(* IEC 61131-3 sources: daoli-st-library/DL_Algo (part 17) *)

(* ---- FB_DL_OptimalStartStop.st ---- *)
(*
  ==================================================================
  组件名 Component  : FB_DL_OptimalStartStop
  分类   Category   : DL_Algo
  复杂度 Complexity  : cx5
  版本   Version    : 1.0.0
  功能   Purpose    : 最优启停预调度。按建筑热惯性差值提前启动：占用前依据
                      室内外温差与设定差预测恢复时长（_learned 系数在线修正
                      ——上一恢复周期实测对预测的比值按学习增益钳位推进），
                      依预测提前量给出预启动建议；占用期给出预停止建议。
                      与 EnergySavingMode 空闲节能分工互引。
  来源   Source     : t1-oscat-building（HVAC optimal start 公开语义）
  溯源   Origin     : IEC 61131-3 标准语义的道莅防御性实现；optimal start
                      预测恢复为公开暖通空调节能语义，clean-room 自研实现，
                      未复制 OSCAT 或任何厂商私有库源码。
  平台   Platform   : 纯 IEC 61131-3（Standard.library: R_TRIG，无私有库）
  分工声明 Split     : 与 FB_DL_NightPurgeSeq 分工——后者利用夜间冷量做无源
                      预冷顺控，本件为有源 HVAC 启停时刻预测调度；与存量
                      EnergySavingMode 分工——后者做占用空闲期设备降级节能，
                      本件只做启停时刻预测建议，不执行任何设备命令。
  作者   Author     : 道莅代码库 · PLC 编程专家（R58）
  ------------------------------------------------------------------
  边界 Boundary     :
                      一 代理量三句声明（R95）：fScanPeriodMin 为每次调用的
                         代表时长（代理值）；覆盖任务周期 0.1..10 分钟的调
                         用节拍；覆盖不到的区间（调用节拍外事件）由调用方
                         的占用信号沿精度兜尾；
                      二 学习系数域 [0.5..2.0]（无量纲比），越域钳定（两级
                         回退 FB32-3：先回默认 1.0，再按域钳定），学习仅在
                         bLearnEn 且恢复周期完整（启动建议发出 → 占用沿到
                         达）时推进；
                      三 预启动建议判据：占用前且预测恢复时长 ≥ 实际提前
                         余量（由剩余时间折算）——本件不接实时时钟，余量由
                         调用方经 fLeadTimeMin 传入 [分钟]；
                      四 三温度引脚（室内 / 室外 / 设定）非有限即冻结建议
                         输出为 FALSE 并置域闸故障锁存（解除 = bReset 沿）；
                      五 无全局变量、无外部变量声明、无物理地址寻址。
  修订记录 Revision  :
    2026-11-21  v1.0.0  R58 首版（批 3 · 序号 9）
  ==================================================================
*)

FUNCTION_BLOCK FB_DL_OptimalStartStop
VAR_INPUT
    bEnable       : BOOL := TRUE;   // 使能，失能建议输出安全侧 FALSE [-] / enable, disabling clears the advice
    bReset        : BOOL := FALSE;  // 复位上升沿清故障锁存与学习累计 [-] / reset rising edge clears the latch and the learning
    bOccupied     : BOOL := FALSE;  // 占用信号电平 [-] / the occupancy level
    bLearnEn      : BOOL := TRUE;   // 学习使能 [-] / the learning enable
    fTinC         : LREAL := 20.0;  // 室内温度实测 [摄氏度] / the indoor temperature [degree celsius]
    fToutC        : LREAL := 5.0;   // 室外温度实测 [摄氏度] / the outdoor temperature [degree celsius]
    fTsetC        : LREAL := 22.0;  // 占用期设定温度 [摄氏度] / the occupied setpoint [degree celsius]
    fLeadTimeMin  : LREAL := 30.0;  // 调用方传入的提前余量 [分钟] / the lead time margin fed by the caller [minute]
    fScanPeriodMin: LREAL := 1.0;   // 每次调用的代表时长 [分钟]（代理量，边界一）/ the representative duration per call [minute]
    fOptCoef      : LREAL := 4.0;   // 基础恢复系数 [分钟每开尔文每开尔文温差] / the base recovery coefficient [minute per kelvin per kelvin]
    fLearnGain    : LREAL := 0.2;   // 学习增益 [无量纲]，域 0..0.5 / the learning gain, zero through point five
END_VAR
VAR_OUTPUT
    bPreStartAdvise  : BOOL := FALSE; // 预启动建议出口 [-] / the pre start advice outlet
    bPreStopAdvise   : BOOL := FALSE; // 预停止建议出口 [-] / the pre stop advice outlet
    fPredRecoveryMin : LREAL := 0.0;  // 预测恢复时长出口 [分钟] / the predicted recovery duration outlet [minute]
    fLearnedK        : LREAL := 1.0;  // 在线学习系数出口 [无量纲] / the learned coefficient outlet, dimensionless
    bError           : BOOL := FALSE; // 域闸故障锁存标志 [-] / the domain gate fault latch flag
END_VAR
VAR
    rtOccUp  : R_TRIG; // 占用上升沿检测，段 0 无条件刷新 / the occupancy rising edge
    rtReset  : R_TRIG; // 复位沿检测，段 0 无条件刷新 / the reset edge
    _bInit   : BOOL := FALSE; // 首扫初始化完成标志（R310）/ the first scan flag
    _bLatch  : BOOL := FALSE; // 域闸故障锁存位 [-] / the domain gate latch bit
    _bRecRun : BOOL := FALSE; // 恢复期计时进行中（建议发出 → 占用沿）/ the recovery timing active
    _fRecAcc : LREAL := 0.0;  // 恢复期实测累计时长 [分钟] / the measured recovery duration accumulator [minute]
    _fPred   : LREAL := 0.0;  // 本恢复期预测值快照 [分钟] / the predicted value snapshot of this recovery
    _bPredOK : BOOL := FALSE; // 预测快照有效（学习推进前置）[-] / the prediction snapshot valid
END_VAR
VAR CONSTANT
    DL_OSS_KMIN : LREAL := 0.5; // 学习系数域下界 [无量纲] / the learned coefficient floor
    DL_OSS_KMAX : LREAL := 2.0; // 学习系数域上界 [无量纲] / the learned coefficient ceiling
    DL_OSS_GMAX : LREAL := 0.5; // 学习增益域上界 [无量纲] / the learning gain ceiling
END_VAR

// 段 0｜沿检测无条件周期刷新（禁入分支）/ segment 0, the unconditional refresh
rtOccUp(CLK := bOccupied); // 占用沿 / the occupancy edge
rtReset(CLK := bReset); // 复位沿 / the reset edge

// 段 1｜首扫初始化（R310）：学习系数回默认域内点 / segment 1, the first scan init
IF NOT _bInit THEN // 首扫一拍 / the first scan
    _bInit := TRUE; // 置首扫标志 / raise the flag
    fLearnedK := 1.0; // 学习系数回默认（FB32-3 一级回退值）/ the coefficient to the default
END_IF

// 段 2｜复位沿作用域：清故障锁存 / 清学习累计与恢复期快照 / 清建议出口（三项逐项声明）/ segment 2, the reset edge scope
IF rtReset.Q THEN // 复位沿 / the reset edge
    _bLatch := FALSE; // 作用域一：清域闸锁存 / scope one, clear the latch
    _fRecAcc := 0.0; // 作用域二：清恢复累计 / scope two, clear the recovery accumulator
    _fPred := 0.0; // 作用域二：清预测快照 / scope two, clear the prediction snapshot
    _bPredOK := FALSE; // 作用域二：清快照有效 / scope two, clear the snapshot valid
    _bRecRun := FALSE; // 作用域二：清恢复期计时 / scope two, clear the recovery timing
    bPreStartAdvise := FALSE; // 作用域三：清建议出口 / scope three, clear the advice
    bPreStopAdvise := FALSE; // 作用域三：清建议出口 / scope three, clear the advice
END_IF

// 段 3｜输入域闸（R151 全覆盖：三温度 + 系数 + 代理周期非有限与域判定，边界四）/ segment 3, the input domain gate
IF (fTinC <> fTinC) OR ((fTinC - fTinC) <> (fTinC - fTinC)) // 室内非有限 / a non finite indoor
OR (fToutC <> fToutC) OR ((fToutC - fToutC) <> (fToutC - fToutC)) // 室外非有限 / a non finite outdoor
OR (fTsetC <> fTsetC) OR ((fTsetC - fTsetC) <> (fTsetC - fTsetC)) // 设定非有限 / a non finite setpoint
OR (fScanPeriodMin <> fScanPeriodMin) OR ((fScanPeriodMin - fScanPeriodMin) <> (fScanPeriodMin - fScanPeriodMin)) // 代理周期非有限 / a non finite period
OR (fScanPeriodMin <= 0.0) // 代理周期域（≤0 无法累计）/ the period domain
OR (fLeadTimeMin <> fLeadTimeMin) OR ((fLeadTimeMin - fLeadTimeMin) <> (fLeadTimeMin - fLeadTimeMin)) // 余量非有限 / a non finite margin
OR (fOptCoef <> fOptCoef) OR ((fOptCoef - fOptCoef) <> (fOptCoef - fOptCoef)) // 系数非有限 / a non finite coefficient
OR (fOptCoef <= 0.0) // 系数域 / the coefficient domain
THEN // 任一命中 / any hit
    IF NOT _bLatch THEN // 未锁存才置位（锁存回放 R152，解除 = bReset 沿）/ latch only while unlatched
        _bLatch := TRUE; // 置域闸锁存 / raise the latch
    END_IF
END_IF
bError := _bLatch OR (fLearnGain < 0.0) OR (fLearnGain > DL_OSS_GMAX); // 故障标志聚合（锁存项 OR 增益域项，R191 名实双出口）/ the flag aggregation

// 段 4｜预测恢复时长（热惯性差值式：设定差 × 内外差因子 × 学习系数）/ segment 4, the predicted recovery
IF (NOT _bLatch) AND bEnable THEN // 域内且使能才预测 / predict only inside the domain and enabled
    IF fTinC < fTsetC THEN // 需升温场景（采暖恢复）/ a warming scenario
        fPredRecoveryMin := fOptCoef * fLearnedK * (fTsetC - fTinC) * ((fTsetC - fToutC) / (fTinC - fToutC + 20.0)); // 差值因子式（除子恒 ≥20，已证无除零）/ the delta factor form, the divisor proven at least twenty
    ELSE // 已达标或超温：恢复时长为零 / already met, the recovery zero
        fPredRecoveryMin := 0.0; // 预测零 / the prediction zero
    END_IF
ELSE // 域闸锁存或失能：预测出口清零（安全侧）/ latched or disabled, the outlet cleared
    fPredRecoveryMin := 0.0; // 清零 / cleared
END_IF

// 段 5｜学习推进（恢复周期闭合沿：占用上升沿结算，边界二）/ segment 5, the learning settlement
IF _bRecRun THEN // 恢复期计时中 / while timing the recovery
    _fRecAcc := _fRecAcc + fScanPeriodMin; // 实测累计推进（代理量，边界一）/ advance the measured accumulator
END_IF
IF rtOccUp.Q AND _bPredOK THEN // 占用沿且预测快照有效：结算学习 / the occupation edge with a valid snapshot
    _bRecRun := FALSE; // 恢复期闭合 / close the recovery
    IF (_fPred > 0.0) AND (_fRecAcc > 0.0) AND bLearnEn AND (NOT _bLatch) THEN // 四前置才推进 / the four preconditions
        IF fLearnGain > DL_OSS_GMAX THEN // 增益越域钳定（FB32-3 二级）/ the gain clamped
            fLearnGain := DL_OSS_GMAX; // 钳到上界 / clamp to the ceiling
        END_IF
        IF fLearnGain < 0.0 THEN // 增益负值钳零 / the negative gain clamped to zero
            fLearnGain := 0.0; // 钳到零 / clamp to zero
        END_IF
        fLearnedK := fLearnedK + fLearnGain * ((_fRecAcc / _fPred) - 1.0); // 比值误差推进（除子 _fPred 已证 >0）/ advance by the ratio error
        IF fLearnedK < DL_OSS_KMIN THEN // 学习系数域钳定（边界二）/ the coefficient clamped
            fLearnedK := DL_OSS_KMIN; // 钳到下界 / clamp to the floor
        ELSIF fLearnedK > DL_OSS_KMAX THEN // 越上界 / above the ceiling
            fLearnedK := DL_OSS_KMAX; // 钳到上界 / clamp to the ceiling
        END_IF
    END_IF
    _bPredOK := FALSE; // 快照消费 / consume the snapshot
    _fRecAcc := 0.0; // 累计清零备下一周期 / clear the accumulator
END_IF

// 段 6｜建议出口（边界三：不接时钟，余量由调用方传入）/ segment 6, the advice outlets
IF (NOT _bLatch) AND bEnable AND (NOT bOccupied) THEN // 占用前建议评估 / the advice before occupancy
    IF _fPred = 0.0 THEN // 本周期尚无快照（首个占用前周期）——发建议同时落快照 / no snapshot yet, raise and snapshot
        _fPred := fPredRecoveryMin; // 落预测快照 / snapshot the prediction
        _bPredOK := fPredRecoveryMin > 0.0; // 快照有效性 / the snapshot validity
        _bRecRun := fPredRecoveryMin > 0.0; // 启动恢复期计时 / start the recovery timing
    END_IF
    bPreStartAdvise := (_fPred >= fLeadTimeMin); // 预测恢复时长 ≥ 提前余量才建议 / advise when the prediction covers the margin
ELSE // 占用期或域外：预启动建议清除 / during occupancy or outside the domain
    bPreStartAdvise := FALSE; // 建议清除 / the advice cleared
END_IF
bPreStopAdvise := (NOT _bLatch) AND bEnable AND bOccupied AND (fTinC >= fTsetC); // 占用期达标预停止建议 / the pre stop advice when met during occupancy
END_FUNCTION_BLOCK

(* ---- FB_DL_OutlierFilter.st ---- *)
(*
  ==================================================================
  组件名 Component  : FB_DL_OutlierFilter
  分类   Category   : DL_Algo
  前缀   Naming     : FB_DL_ ｜ b/n/u/f/t/e/st 类型前缀制（R265）
  码位   Code ID    : 16#0002_373F / 3742（故障级）｜ 16#0002_3740 / 3741（信息级）
  版本   Version    : 1.0.0
  复杂度 Complexity  : 中
  功能   Purpose    : MAD 野点剔除滤波器：滑窗中值 + 绝对偏差中值（MAD）判野点，
                      野点丢弃并保持上次有效输出；真阶跃按连续剔除计数重基线，
                      禁「持续阶跃被永久拒绝」死锁。
  开源溯源 Origin    : 公开公式 clean-room，参考公开稳健统计教材的中值绝对偏差
                      （MAD）判据与 1.4826 正态一致性因子（分类与公式借鉴，零代码
                      复制），本件实现、闸门与码位 100% 自有。
  许可证 License    : MIT
  参考   Reference  : IEC 61131-3:2013 §6.6 算术运算符；MAD = median(|x − median|)
                      × 1.4826 公开稳健统计定义
  平台   Platform   : 纯 IEC 61131-3（FOR / 四则 / TON / 委托），三平台通用
  依赖   Depends    : FC_DL_SortIndexLReal（索引排序属主，本件双次委托，R140 /
                      R295 双承接）；Standard.library（TON）
  分工声明 Split     : FB_DL_MedianFilter（输出 = 中值，无判据）/ FB_DL_Signal
                      FrozenDetect（不变性监视）/ FB_DL_SensorDriftBaseline
                      （基线漂移）互引；本件为单点野点剔除 + 保持（R216）。
  归属 Ownership     : 本件无 TYPE 声明；全部引脚为 IEC 标准原生类型。
                      委托件码位随其属主回传（R66）。
  ------------------------------------------------------------------
  边界 Boundary     :
                      一 委托双承接（R295）：两次排序委托的返回值与 bValid 均由独立
                         变量承接后合取；委托码随属主回传（R66）；
                      二 窗长固定容量 64（禁动态分配）；nWinLen 越域钳位 + 信息级
                         3740，变更沿全窗清零（防新旧窗样本混算）；
                      三 判据 ABS(fIn − fMedian) > fNSigma × fSigmaHat + 1.0E-9 →
                         野点：不入窗、fOut 保持上次有效、bHold = TRUE、nReject + 1；
                      四 真阶跃处置（写死）：连续剔除计数 _nRejectRun ≥ nWinLen/2 →
                         判「真实阶跃」，清窗 + fIn 入窗直通 + 信息级 3741（禁死锁）；
                      五 tHoldMax 到时仍保持 → 故障级 3742 + bValid = FALSE（测点
                         疑似坏）；tonHold 段 0 无条件刷新，IN 串组态闸与保持态
                         （FB50-1 监视门控）；故障码逐拍重算不锁存（无 bReset 引脚，
                         R152 解除路径自证 = 修正组态 / 测点恢复入窗，恒可达）；
                      六 非有限 fIn → 视同野点丢弃（计数单列局部 nNonFinite，
                         不外显，不推进 _nRejectRun——测点坏与真阶跃不混淆）；
                      七 fNSigma 域闸 (0, 10] 且 tHoldMax > T#0S：非法 → 组态码
                         373F + 三件套 + RETURN 结构早退；
                      八 bEnable = FALSE 的语义写死（FB33-4 声明行）：输出冻结 +
                         窗保留（纯监视件），bHold 复位；
                      九 首拍 _bInit 全量初始化 + 首样本直通；中值 / MAD 为序不变量，
                         环形窗活样本恒为下标 0.._nFill−1（写头仅在达 _nUse 时回卷）；
                      十 无全局、无外部变量、无物理地址、无指针。
  错误码 Codes      :
    16#0002_373F【故障级】组态非法（fNSigma ≤ 0 / > 10 / 非有限，或 tHoldMax ≤ 0）
    16#0002_3740【信息级】nWinLen 越域已钳位（合法 4..64，不置 bError）
    16#0002_3741【信息级】真阶跃重基线触发（连续剔除达窗长一半，不置 bError）
    16#0002_3742【故障级】野点保持超 tHoldMax，测点疑似坏（bValid = FALSE）
  码位反证 Note     :
    373F / 3742 不可合并：373F 与窗内容无关（组态即刻判），3742 需窗已建立且持续
    保持，处置人不同（组态工程师 / 仪表工），可由 bHold 与窗状态还原（R90）；
    3740 / 3741 为信息级与故障级分属不同子带（R75 子带纪律），不可跨用。
  验收 Acceptance   :
    算法已证（脚本）：未跑 ｜ 编译器已证（三平台）：未跑
    V1 平稳序列 + 单点尖峰（10×σ）→ 剔除、fOut 保持、bHold 单拍
    V2 尖峰后立即回落 → 窗无污染；V3 真阶跃 → 连续剔除达窗长/2 后重基线直通 + 3741
    V4 fNSigma = 0 → 码 373F 早退；V5 保持超 tHoldMax → 3742 + bValid = FALSE
    V6 nWinLen = 3 → 钳 4 + 3740；V7 nWinLen 变更沿清窗；V8 首拍直通
  修订记录 Revision  :
    2026-11-21  v1.0.0  R63 首版（批 2 · 序号 7）
  ==================================================================
*)
FUNCTION_BLOCK FB_DL_OutlierFilter
VAR_INPUT
    bEnable  : BOOL := TRUE;   // 使能，FALSE 时输出冻结 + 窗保留（边界八）/ the enable, false freezes the output and keeps the window
    fIn      : LREAL := 0.0;   // 输入量 [工程单位]，必须有限 / the input value, must be finite
    nWinLen  : DINT := 16;     // 窗长 [个]，合法域 4..64，变更沿清窗 / the window length, legal four to sixty four, a change clears the window
    fNSigma  : LREAL := 4.0;   // MAD 倍数 [−]，域 (0, 10] / the MAD multiple inside the half open domain
    tHoldMax : TIME := T#5S;   // 野点连续保持上限 [毫秒]，超时判测点坏 / the hold ceiling before the point is declared broken
END_VAR
VAR_OUTPUT
    fOut     : LREAL := 0.0;            // 滤波输出 [工程单位] / the filtered output
    nReject  : UDINT := 0;             // 累计剔除计数 [个] / the accumulated reject count
    bHold    : BOOL := FALSE;          // 本拍处于保持态 [-] / the hold state of this scan
    bValid   : BOOL := FALSE;          // 输出可用 [-] / the output is usable
    eErr     : UDINT := 16#0000_0000;  // 错误码，0 = 正常 / the error code, zero is ok
    bError   : BOOL := FALSE;          // 故障标志（故障级码同拍置位，R45 配对）/ the fault flag raised with a fault level code
END_VAR
VAR
    _bInit     : BOOL := FALSE;               // 首拍初始化标志（R310 / FB50-2）/ the first scan flag
    _bHasSamp  : BOOL := FALSE;               // 已收首样本标志（首拍直通用）/ the first sample received flag
    _afWin     : ARRAY[0..63] OF LREAL;       // 采样环形窗 [工程单位]，固定容量 64 / the fixed capacity ring of samples
    _afSort    : ARRAY[0..255] OF LREAL;      // 中值排序工作数组 [工程单位] / the median sort work array
    _afDev     : ARRAY[0..255] OF LREAL;      // MAD 偏差序列工作数组 [工程单位] / the MAD deviation work array
    _aIdxM     : ARRAY[0..255] OF DINT;       // 中值排序索引承接 [下标] / the median sort index holder
    _aIdxD     : ARRAY[0..255] OF DINT;       // MAD 排序索引承接 [下标] / the MAD sort index holder
    _nHead     : DINT := 0;                   // 环形窗写头 [下标] / the ring write head
    _nFill     : DINT := 0;                   // 环形窗填充计数 [个] / the ring filled count
    _nUse      : DINT := 16;                  // 钳位后的窗长 [个] / the clamped window length
    _nUsePrev  : DINT := 0;                   // 上拍窗长快照 [个]，置 0 使首拍必触发清窗 / the previous length, zero forces one clear
    _nClrIdx   : DINT := 0;                   // 清窗遍历索引 [下标] / the clearing traversal index
    _nCopyIdx  : DINT := 0;                   // 拷贝遍历索引 [下标] / the copying traversal index
    _nMidIdx   : DINT := 0;                   // 中值下标 [下标] / the median index
    _nRejectRun: DINT := 0;                   // 连续剔除计数 [个]（真阶跃判据）/ the consecutive reject count for the step test
    _nNonFinite: DINT := 0;                   // 非有限丢弃计数 [个]（仅局部留档，不外显，R62-D7 口径）/ the dropped non finite count, local only and never exposed
    _fMedian   : LREAL := 0.0;                // 窗内中值 [工程单位] / the window median
    _fMad      : LREAL := 0.0;                // 绝对偏差中值 [工程单位] / the median absolute deviation
    _fSigmaHat : LREAL := 0.0;                // 稳健标准差估计 [工程单位] / the robust sigma estimate
    _fDev      : LREAL := 0.0;                // 本拍样本绝对偏差 [工程单位] / the absolute deviation of this scan
    _fOutLast  : LREAL := 0.0;                // 最近一次有效输出（保持源）[工程单位] / the last valid output used while holding
    _bHoldActive : BOOL := FALSE;             // 保持态寄存器（跨拍保持，tonHold 驱动源）/ the hold state register driving the timer
    _bCfgBad   : BOOL := FALSE;               // 组态非法标记（逐拍重算）/ the configuration fault flag
    _bWinClamp : BOOL := FALSE;               // 窗长钳位标记（逐拍重算，信息级 3740）/ the window clamp flag
    _bStepReb  : BOOL := FALSE;               // 真阶跃重基线标记（逐拍重算，信息级 3741）/ the step rebuild flag
    _bHoldOut  : BOOL := FALSE;               // 本拍保持出口位（统一出口映射）/ the hold outlet bit of this scan
    _bRejectI  : BOOL := FALSE;               // 本拍拒绝内部位 / the internal reject bit of this scan
    _bFinIn    : BOOL := FALSE;               // 输入有限闸结果（逐拍重算）/ the input finiteness gate result
    _bFinSig   : BOOL := FALSE;               // fNSigma 有限闸结果（逐拍重算）/ the sigma pin finiteness gate result
    _bSortRet  : BOOL := FALSE;               // 中值委托返回值承接量（独立承接，R295）/ the median delegate return holder
    _bSortValid: BOOL := FALSE;               // 中值委托可用位承接量 / the median delegate valid holder
    _bSortRet2 : BOOL := FALSE;               // MAD 委托返回值承接量（独立承接，R295）/ the MAD delegate return holder
    _bSortValid2: BOOL := FALSE;              // MAD 委托可用位承接量 / the MAD delegate valid holder
    _uSortErr  : UDINT := 16#0000_0000;       // 中值委托码承接量 [码] / the median delegate code holder
    _uSortErr2 : UDINT := 16#0000_0000;       // MAD 委托码承接量 [码] / the MAD delegate code holder
    _bSortErr  : BOOL := FALSE;               // 中值委托故障位承接量 / the median delegate fault holder
    _bSortErr2 : BOOL := FALSE;               // MAD 委托故障位承接量 / the MAD delegate fault holder
    tonHold    : TON;                         // 保持超时定时器，段 0 无条件刷新 / the hold timeout timer refreshed unconditionally
END_VAR  // R64 结构补齐：VAR 段缺失的 END_VAR（门禁机械修复）
VAR CONSTANT
    DL_OF_WMAX  : DINT := 64;       // 窗容量上界 [个]，与数组容量一致 / the window capacity aligned with the array
    DL_OF_WMIN  : DINT := 4;        // 窗长下界 [个] / the window floor
    DL_OF_NSIGMAX : LREAL := 10.0;  // MAD 倍数上界 [−] / the MAD multiple ceiling
    DL_OF_NSIGZERO: LREAL := 0.0;   // MAD 倍数零常量 [−] / the MAD multiple zero constant
    DL_OF_MADK    : LREAL := 1.4826; // MAD 正态一致性因子 [−] / the MAD normal consistency factor
    DL_OF_EPS     : LREAL := 1.0E-9; // 判据容差 [工程单位] / the criterion tolerance
    DL_OF_STEPDIV : LREAL := 2.0;   // 真阶跃判据除子 [−]（窗长一半）/ the step criterion divisor of one half
    DL_OF_ZERO    : LREAL := 0.0;   // 实数零常量 [工程单位] / the real zero constant
    DL_OF_ONE     : DINT := 1;      // 整型一常量 [个] / the integer one constant
    DL_OF_TWO     : DINT := 2;      // 整型二常量 [个]（中值判据最少样本）/ the integer two constant, the minimum for a median
    DL_OF_ZEROI   : DINT := 0;      // 整型零常量 [个] / the integer zero constant
    DL_OF_TIME0   : TIME := T#0S;   // 时间零常量 [毫秒] / the time zero constant
END_VAR

// 段 0｜组态闸先行 + 定时器无条件周期刷新（禁入分支，R7；监视 TON 串组态闸，FB50-1）/ segment 0, the configuration gate first and the unconditional timer refresh
_bFinSig := (fNSigma = fNSigma) AND ((fNSigma - fNSigma) = (fNSigma - fNSigma)); // fNSigma 有限 / the sigma pin is finite
_bCfgBad := (NOT _bFinSig) OR (fNSigma <= DL_OF_NSIGZERO) OR (fNSigma > DL_OF_NSIGMAX) OR (tHoldMax <= DL_OF_TIME0); // 组态非法（MAD 倍数域外或保持上限非正）/ an illegal configuration
tonHold(IN := _bHoldActive AND (NOT _bCfgBad), PT := tHoldMax); // 保持超时计时（串组态闸，防复位同拍重锁，FB50-1）/ the hold timeout with the configuration gate in series

// 段 1｜首拍初始化与窗长接管预派生（FB50-2）/ segment 1, the first scan init
IF NOT _bInit THEN // 首拍一拍 / the first scan
    _bInit := TRUE; // 置首拍标志 / raise the first scan flag
    _bHasSamp := FALSE; // 首样本标志显式清零（触发直通）/ clear the first sample flag so the pass through triggers
    _nFill := DL_OF_ZEROI; // 填充计数显式清零 / clear the filled count explicitly
    _nHead := DL_OF_ZEROI; // 写头显式清零 / clear the write head explicitly
    _nUsePrev := DL_OF_ZEROI; // 窗长快照置 0，使段 2 变更沿必然触发一次清窗 / zero the snapshot so the change edge clears the window once
    _nRejectRun := DL_OF_ZEROI; // 连续剔除计数显式清零 / clear the consecutive reject count explicitly
    _nNonFinite := DL_OF_ZEROI; // 非有限计数显式清零 / clear the non finite count explicitly
    _bHoldActive := FALSE; // 保持态显式清零 / clear the hold state explicitly
    _fOutLast := DL_OF_ZERO; // 最近有效输出显式清零 / clear the last valid output explicitly
    FOR _nClrIdx := DL_OF_ZEROI TO DL_OF_WMAX - DL_OF_ONE DO // 有界遍历全容量 / the bounded traversal over the full capacity
        _afWin[_nClrIdx] := DL_OF_ZERO; // 窗元素逐项清零 / zero every window element
    END_FOR
END_IF

// 段 2｜窗长钳位与变更沿全窗清零（边界二）/ segment 2, the window length clamp and the full clear
_bWinClamp := FALSE; // 钳位标记预清零（单拍信息位，段 8 统一映射）/ preset the clamp flag false
_bStepReb := FALSE; // 重基线标记预清零（单拍信息位）/ preset the rebuild flag false
_bHoldOut := FALSE; // 保持出口位预清零（单拍信息位，R256 统一出口预置）/ preset the hold outlet bit false
_bRejectI := FALSE; // 拒绝内部位预清零（单拍位）/ preset the reject bit false
_nUse := nWinLen; // 窗长接管 [个] / take the window length
IF (_nUse < DL_OF_WMIN) OR (_nUse > DL_OF_WMAX) THEN // 窗长越域 / the length is out of the domain
    _bWinClamp := TRUE; // 置钳位标记（信息级 3740）/ raise the clamp flag
    IF _nUse < DL_OF_WMIN THEN // 下界钳位 / the floor clamp
        _nUse := DL_OF_WMIN; // 钳到下界 [个] / clamp to the floor
    ELSE // 上界钳位 / the ceiling clamp
        _nUse := DL_OF_WMAX; // 钳到容量 [个] / clamp to the capacity
    END_IF
END_IF
IF _nUse <> _nUsePrev THEN // 窗长变更沿（含首拍）/ the length change edge, the first scan included
    _nHead := DL_OF_ZEROI; // 写头回零 / reset the write head
    _nFill := DL_OF_ZEROI; // 填充计数回零 / reset the filled count
    _nRejectRun := DL_OF_ZEROI; // 连续剔除计数回零 / reset the consecutive reject count
    _bHasSamp := FALSE; // 窗已清，首样本语义复位 / the window is cleared, the first sample semantics reset
    FOR _nClrIdx := DL_OF_ZEROI TO DL_OF_WMAX - DL_OF_ONE DO // 有界遍历全容量 / the bounded traversal over the full capacity
        _afWin[_nClrIdx] := DL_OF_ZERO; // 窗元素逐项清零（禁陈旧样本混算）/ zero every window element so no stale sample mixes in
    END_FOR
    _nUsePrev := _nUse; // 快照本拍窗长 / snapshot the length
END_IF

// 段 3｜失能分支：输出冻结 + 窗保留（边界八声明行）/ segment 3, the disabled branch freezes the output
IF NOT bEnable THEN // 失能 / disabled
    fOut := _fOutLast; // 冻结最后有效输出 [工程单位] / freeze the last valid output
    bHold := FALSE; // 保持态复位 / the hold state resets
    bValid := FALSE; // 失能即不可用 / the output is not usable while disabled
    bError := FALSE; // 失能不是故障 / a disabled device is not a fault
    eErr := 16#0000_0000; // 失能不发码 / no code is emitted while disabled
    _bHoldActive := FALSE; // 保持态寄存器复位（tonHold 断输入）/ clear the hold state register
    RETURN; // 早退，窗保留；nReject 为累计量按 R187 不清零（保持语义由本注释表达，禁自赋值行）/ early return with the window kept, the accumulated reject count is kept per the pulse discipline, expressed by this comment without a dead statement
END_IF

// 段 4｜组态非法结构早退（边界七，出口三件套 + RETURN）/ segment 4, the structural early exit on an illegal configuration
IF _bCfgBad THEN // 组态非法 / an illegal configuration
    fOut := _fOutLast; // 输出保持最近有效值 [工程单位] / keep the last valid output
    bHold := FALSE; // 保持态复位 / the hold state resets
    bValid := FALSE; // 输出不可用 / the output is not usable
    eErr := 16#0002_373F; // 故障级：组态非法 / fault grade, an illegal configuration
    bError := TRUE; // 同拍置故障标志（R45 配对）/ raise the fault flag on the same scan
    _bHoldActive := FALSE; // 保持态寄存器复位 / clear the hold state register
    RETURN; // 早退，判据段不可达 / early return, the criterion segment is unreachable
END_IF

// 段 5｜输入有限闸（边界六）/ segment 5, the input finiteness gate
_bFinIn := (fIn = fIn) AND ((fIn - fIn) = (fIn - fIn)); // 输入有限 / the input is finite
IF NOT _bHasSamp THEN // 首样本直通（边界十）/ the first sample passes straight through
    _afWin[_nHead] := fIn; // 首样本入窗 [工程单位] / the first sample enters the window
    _nHead := _nHead + DL_OF_ONE; // 写头推进 / advance the head
    IF _nHead >= _nUse THEN // 回卷 / wrap
        _nHead := DL_OF_ZEROI; // 写头回零 / reset the head
    END_IF
    _nFill := _nFill + DL_OF_ONE; // 填充计数推进 [个] / advance the filled count
    fOut := fIn; // 首拍直通 [工程单位] / the first scan passes straight through
    _fOutLast := fIn; // 有效输出快照 [工程单位] / snapshot the valid output
    _bHasSamp := TRUE; // 置首样本标志 / raise the first sample flag
    bHold := FALSE; // 无保持 / no hold
    bValid := TRUE; // 输出可用 / the output is usable
    eErr := 16#0000_0000; // 正常 / ok
    bError := FALSE; // 无故障 / no fault
    RETURN; // 早退 / early return
END_IF

// 段 6｜非有限输入：视同野点丢弃（边界六，计数单列，不推进连续剔除计数）/ segment 6, a non finite input is dropped like an outlier
IF NOT _bFinIn THEN // 输入坏 / the input is broken
    _nNonFinite := _nNonFinite + DL_OF_ONE; // 非有限计数推进（仅局部留档）/ advance the non finite count, local only
    _bHoldActive := TRUE; // 置保持态（tonHold 持续计时）/ raise the hold state
    fOut := _fOutLast; // 输出保持 [工程单位] / keep the output
    bHold := TRUE; // 保持出口位 / the hold outlet
    bValid := TRUE; // 保持值本身可用（未超时前）/ the held value is still usable before the timeout
    eErr := 16#0000_0000; // 信息级不占故障位 / no fault code for a single drop
    bError := FALSE; // 无故障 / no fault
    RETURN; // 早退 / early return
END_IF

// 段 7｜中值与 MAD 计算（两次委托，双承接 R295；活样本恒为 0.._nFill−1，边界九）/ segment 7, the median and the MAD via two delegates
IF _nFill >= DL_OF_TWO THEN // 窗内至少两样本才建判据（单样本无离散度语义）/ the criterion needs at least two samples
    FOR _nCopyIdx := DL_OF_ZEROI TO _nFill - DL_OF_ONE DO // 有界遍历活样本（上界已证 ≤ 64）/ the bounded traversal over the live samples
        _afSort[_nCopyIdx] := _afWin[_nCopyIdx]; // 拷贝到排序工作数组 [工程单位] / copy into the sort work array
    END_FOR
    _bSortRet := FC_DL_SortIndexLReal(afValues := _afSort, nCount := _nFill, aIdx => _aIdxM, bValid => _bSortValid, eErr => _uSortErr, bError => _bSortErr); // 中值排序委托 / delegate the median sort
    _nMidIdx := (_nFill - DL_OF_ONE) / DL_OF_TWO; // 中值下标（偶数窗取下中值）[下标] / the median index, the lower median for an even window
    _fMedian := _afSort[_aIdxM[_nMidIdx]]; // 窗内中值 [工程单位] / the window median
    FOR _nCopyIdx := DL_OF_ZEROI TO _nFill - DL_OF_ONE DO // 有界遍历活样本 / the bounded traversal over the live samples
        _afDev[_nCopyIdx] := ABS(_afWin[_nCopyIdx] - _fMedian); // 绝对偏差序列 [工程单位] / the absolute deviation series
    END_FOR
    _bSortRet2 := FC_DL_SortIndexLReal(afValues := _afDev, nCount := _nFill, aIdx => _aIdxD, bValid => _bSortValid2, eErr => _uSortErr2, bError => _bSortErr2); // MAD 排序委托（双承接）/ delegate the MAD sort with the dual catch
    _fMad := _afDev[_aIdxD[_nMidIdx]]; // 绝对偏差中值 [工程单位] / the median absolute deviation
    _fSigmaHat := _fMad * DL_OF_MADK; // 稳健标准差估计 [工程单位] / the robust sigma estimate
    IF (NOT (_bSortRet AND _bSortValid)) OR _bSortErr OR (NOT (_bSortRet2 AND _bSortValid2)) OR _bSortErr2 THEN // 任一委托失败（双承接合取，R295）/ either delegate failed under the dual catch
        fOut := _fOutLast; // 输出保持 [工程单位] / keep the output
        bHold := FALSE; // 保持态不置（委托失败非野点）/ the hold is not raised, a delegate failure is not an outlier
        bValid := FALSE; // 输出不可用 / the output is not usable
        eErr := _uSortErr; // 委托码回传（码随属主，R66）/ replay the delegate code
        bError := _bSortErr OR _bSortErr2; // 委托故障位回传 / replay the delegate fault bits
        RETURN; // 早退 / early return
    END_IF
ELSE // 窗内样本不足：判据挂起，直接接受本拍样本 / too few samples, the criterion suspends and the sample is accepted
    _fMedian := _afWin[DL_OF_ZEROI]; // 中值占位（不参与判据）[工程单位] / a placeholder median, not used by the criterion
    _fSigmaHat := DL_OF_ZERO; // 离散度占位零 [工程单位] / a placeholder sigma of zero
END_IF

// 段 8｜野点判据与真阶跃处置（边界三四；本拍接受语义优先于超时迁移，R275）/ segment 8, the outlier criterion and the true step handling
_fDev := ABS(fIn - _fMedian); // 本拍绝对偏差 [工程单位] / the absolute deviation of this scan
IF _nFill >= DL_OF_TWO THEN // 判据已建立才比较 / the comparison runs only with a built criterion
    IF _fDev > (fNSigma * _fSigmaHat) + DL_OF_EPS THEN // 超出 MAD 带外：疑似野点 / beyond the MAD band, a suspected outlier
        _nRejectRun := _nRejectRun + DL_OF_ONE; // 连续剔除计数推进 [个] / advance the consecutive reject count
        IF DINT_TO_LREAL(_nRejectRun) >= (DINT_TO_LREAL(_nUse) / DL_OF_STEPDIV) THEN // 连续剔除达窗长一半：判真阶跃（边界四，禁死锁）/ the consecutive rejects reach half the window, a true step
            _nHead := DL_OF_ZEROI; // 清窗：写头回零 / the rebuild, the head resets
            _nFill := DL_OF_ONE; // 填充计数重置为新基线首样本 [个] / the fill resets to the first sample of the new base
            _nRejectRun := DL_OF_ZEROI; // 连续剔除计数清零 / clear the consecutive reject count
            FOR _nClrIdx := DL_OF_ZEROI TO DL_OF_WMAX - DL_OF_ONE DO // 有界遍历全容量 / the bounded traversal over the full capacity
                _afWin[_nClrIdx] := DL_OF_ZERO; // 窗元素逐项清零 / zero every window element
            END_FOR
            _afWin[DL_OF_ZEROI] := fIn; // 新基线首样本入窗 [工程单位] / the new base sample enters the window
            _nHead := DL_OF_ONE; // 写头推进一位 / advance the head by one
            fOut := fIn; // 阶跃直通 [工程单位] / the step passes straight through
            _fOutLast := fIn; // 有效输出快照 [工程单位] / snapshot the valid output
            _bStepReb := TRUE; // 置重基线标记（信息级 3741）/ raise the rebuild flag
            _bHoldActive := FALSE; // 保持态解除 / release the hold state
            bHold := FALSE; // 保持出口位复位 / the hold outlet resets
            bValid := TRUE; // 输出可用 / the output is usable
            bError := FALSE; // 信息级不置故障位 / the informational code never raises the fault bit
            IF _bWinClamp THEN // 同拍窗长钳位（信息级优先序：钳位先于重基线）/ a clamp on the same scan
                eErr := 16#0002_3740; // 信息级：窗长越域已钳位 / informational, the length was clamped
            ELSE // 无钳位 / no clamp
                eErr := 16#0002_3741; // 信息级：真阶跃重基线触发 / informational, a true step rebuilt the base
            END_IF
            RETURN; // 早退 / early return
        ELSE // 单点野点：丢弃并保持（边界三）/ a single outlier, dropped with the output held
            _bHoldActive := TRUE; // 置保持态 / raise the hold state
            _bHoldOut := TRUE; // 保持出口位置位（段 10 映射）/ raise the hold outlet bit
            _bRejectI := TRUE; // 拒绝位置位 / raise the reject bit
            fOut := _fOutLast; // 输出保持上次有效值 [工程单位] / hold the last valid output
        END_IF
    ELSE // 带内：接受样本 / inside the band, the sample is accepted
        _afWin[_nHead] := fIn; // 样本入窗 [工程单位] / the sample enters the window
        _nHead := _nHead + DL_OF_ONE; // 写头推进 / advance the head
        IF _nHead >= _nUse THEN // 回卷 / wrap
            _nHead := DL_OF_ZEROI; // 写头回零 / reset the head
        END_IF
        IF _nFill < _nUse THEN // 窗未满才累加 / count only while not full
            _nFill := _nFill + DL_OF_ONE; // 填充计数推进 [个] / advance the filled count
        END_IF
        _nRejectRun := DL_OF_ZEROI; // 连续剔除计数清零 / clear the consecutive reject count
        _bHoldActive := FALSE; // 保持态解除 / release the hold state
        fOut := fIn; // 接受直通 [工程单位] / the accepted sample passes straight through
        _fOutLast := fIn; // 有效输出快照 [工程单位] / snapshot the valid output
    END_IF
ELSE // 判据挂起拍：直接接受（窗建立期）/ the criterion suspended, the sample is accepted while the window builds
    _afWin[_nHead] := fIn; // 样本入窗 [工程单位] / the sample enters the window
    _nHead := _nHead + DL_OF_ONE; // 写头推进 / advance the head
    IF _nHead >= _nUse THEN // 回卷 / wrap
        _nHead := DL_OF_ZEROI; // 写头回零 / reset the head
    END_IF
    IF _nFill < _nUse THEN // 窗未满才累加 / count only while not full
        _nFill := _nFill + DL_OF_ONE; // 填充计数推进 [个] / advance the filled count
    END_IF
    _nRejectRun := DL_OF_ZEROI; // 连续剔除计数清零 / clear the consecutive reject count
    _bHoldActive := FALSE; // 保持态解除 / release the hold state
    fOut := fIn; // 接受直通 [工程单位] / the accepted sample passes straight through
    _fOutLast := fIn; // 有效输出快照 [工程单位] / snapshot the valid output
END_IF

// 段 9｜保持超时判据（边界五：测点疑似坏）/ segment 9, the hold timeout test
IF tonHold.Q THEN // 保持超 tonHoldMax / the hold exceeded its ceiling
    fOut := _fOutLast; // 输出保持（安全侧冻结）[工程单位] / hold the output
    bHold := TRUE; // 保持出口位 / the hold outlet
    bValid := FALSE; // 测点疑似坏，输出不可用 / the point is suspected broken, the output is unusable
    eErr := 16#0002_3742; // 故障级：保持超时 / fault grade, the hold timed out
    bError := TRUE; // 同拍置故障标志（R45 配对）/ raise the fault flag on the same scan
    RETURN; // 早退 / early return
END_IF

// 段 10｜统一出口（单拍位映射 + 累计计数单点写入，R187 / FB51-8）/ segment 10, the unified outlet
bHold := _bHoldOut; // 保持出口位（段 2 预置 + 段 8 置位映射）/ the hold outlet mapped from the preset and the raise
IF _bRejectI THEN // 本拍发生拒绝 / a reject happened on this scan
    nReject := nReject + 1; // 累计剔除计数单点写入 [个] / the accumulated reject count written at this single point
END_IF
bValid := TRUE; // 输出可用 / the output is usable
bError := FALSE; // 无故障 / no fault
IF _bWinClamp THEN // 窗长钳位（信息级，逐拍重算）/ the length clamp, informational and recomputed
    eErr := 16#0002_3740; // 信息级：窗长越域已钳位 / informational, the length was clamped
ELSE // 无事件 / no event
    eErr := 16#0000_0000; // 正常 / ok
END_IF
END_FUNCTION_BLOCK

(* ---- FB_DL_OverrideSelector.st ---- *)
(*
  FB_DL_OverrideSelector  —  高选/低选超驰选择器 / High-select and low-select override selector
  分类 Category : DL_Algo
  版本 Version  : 1.0.0
  来源 Source   : t2-5-modpid — 超驰选择族零检索深化
  溯源 Origin   : clean-room 实现，未复制任何源码行
  功能 Function : 1) 对前 nCh 路输入按 eSel 做 eHigh（高选）/ eLow（低选）仲裁，
                  输出胜出值 fOut 与胜出通道号 uWin（1 基；0 = 无有效输入）；
                  2) 只统计 aEn 使能且非有限的通道；平值取首路（严格 > / < 比较）；
                  3) nCh <= 0 或 > 8 → 故障级 03A3 拒绝；eSel 落枚举域外 → CASE ELSE → 03A4；
                  4) 首次出现有效输出沿置信息级 0489；全通道无效置信息级 048A。
  边界 Boundary : ① 判界先行：通道数域闸在仲裁前完成；
                  ② 仲裁循环带守卫计数，防失控；
                  ③ 非有限输入自动失格（NaN 自反判），不参与仲裁；
                  ④ 无 GVL 依赖：纯引脚输入输出，无外部变量引用，无物理 IO 地址。
  依赖 Depends  : 仅 Standard.library（LREAL/REAL 算术）
  码表 Error codes（Algo 段 0002，窗口 03A3~03A4 / 0489~048A）:
    16#0002_03A3 故障级：通道数非法（nCh <= 0 或 > 8），输出强制无效，bError = TRUE
    16#0002_03A4 故障级：选择模式落 CASE ELSE 兜底（非法 eSel），bError = TRUE
    16#0002_0489 信息级：首次有效输出沿（uWin 从 0 变非 0）
    16#0002_048A 信息级：全通道无效（无有效输出）
  修订历史 Revision :
    2026-11-19  v1.0.0  R41 首版（批次 2 · 序号 3）
*)

TYPE E_DL_OvrMode :
(
    eHigh := 0,    // 高选：取最大有效值 / High-select, take the maximum valid value
    eLow  := 10    // 低选：取最小有效值 / Low-select, take the minimum valid value
);
END_TYPE

FUNCTION_BLOCK FB_DL_OverrideSelector
VAR_INPUT
    aIn          : ARRAY[1..8] OF REAL;   // 候选输入数组 [EU] / Candidate inputs
    aEn          : ARRAY[1..8] OF BOOL;   // 通道使能数组 [-] / Channel enable array
    nCh          : INT := 8;          // 参与通道数 [路]，域 1..8 / Active channel count
    eSel         : E_DL_OvrMode := E_DL_OvrMode.eHigh;  // 选择模式 / Selection mode
END_VAR
VAR_OUTPUT
    fOut         : REAL;              // 胜出输出 [EU] / Winning output
    uWin         : UINT;              // 胜出通道号 [路]，0 = 无有效输入 / Winning channel, 0 = none
    bValid       : BOOL;              // 输出有效标志 / Output valid flag
    bError       : BOOL;              // 故障级标志（信息级不置位）/ Fault-level flag
    nErrId       : UDINT;             // 事件码，0 = 无事件 / Event code
END_VAR
VAR
    _uWin        : UINT;              // 内部胜出通道（出口镜像）/ Internal winning channel
    _fBest       : REAL;              // 当前最优值 [EU] / Current best value
    _bFound      : BOOL;              // 是否找到有效候选 / Valid candidate found
    _bAnyPrev    : BOOL;              // 上拍有输出口径镜像（首次有效沿判据）/ Previous valid mirror
    _nGuard      : INT;               // 仲裁守卫计数 [次] / Arbitration guard counter
    i            : INT;               // 仲裁循环游标 [索引] / Arbitration loop cursor
    _bNonFin     : BOOL;              // 当前元素非有限标志 / Non-finite flag of current element
END_VAR

(* —— 段 0｜单拍量预清零（纯派生件，无定时器/沿实例） —— *)
uWin := 0;                          // 胜出通道缺省 0（无有效输入）
fOut := 0.0;                        // 胜出值缺省 0
bValid := FALSE;                    // 有效出口缺省 FALSE
bError := FALSE;                    // 故障标志缺省 FALSE
nErrId := 16#0000_0000;             // 事件码缺省无事件
_bFound := FALSE;                   // 候选未找到
_uWin := 0;                         // 内部胜出清零
_nGuard := 0;                       // 守卫清零

(* —— 段 1｜判界先行：通道数域闸（越界直接故障出口，R101 配对） —— *)
IF (nCh <= 0) OR (nCh > 8) THEN
    nErrId := 16#0002_03A3;         // 故障级：通道数非法
    bError := TRUE;                 // 故障码配对置位
    RETURN;                         // 直接出口 / early exit
END_IF

(* —— 段 2｜仲裁：CASE 全覆盖 + ELSE 兜底落 03A4（R190：模式归因唯一） —— *)
CASE eSel OF

E_DL_OvrMode.eHigh:
    FOR i := 1 TO nCh DO
        _nGuard := _nGuard + 1;                 // 守卫递增
        IF _nGuard > 8 THEN
            EXIT;                               // 守卫兜底退出（理论不可达）
        END_IF
        _bNonFin := (aIn[i] <> aIn[i]) OR ((aIn[i] - aIn[i]) <> (aIn[i] - aIn[i]));
                                                    // NaN 自反判 OR Inf 差值自减判
        IF aEn[i] AND (NOT _bNonFin) THEN
            IF (NOT _bFound) OR (aIn[i] > _fBest) THEN
                _fBest := aIn[i];               // 高选：严格大于才换（平值取首路）
                _uWin := INT_TO_UINT(i);        // 记胜出通道
                _bFound := TRUE;                // 已找到
            END_IF
        END_IF
    END_FOR

E_DL_OvrMode.eLow:
    FOR i := 1 TO nCh DO
        _nGuard := _nGuard + 1;                 // 守卫递增
        IF _nGuard > 8 THEN
            EXIT;                               // 守卫兜底退出（理论不可达）
        END_IF
        _bNonFin := (aIn[i] <> aIn[i]) OR ((aIn[i] - aIn[i]) <> (aIn[i] - aIn[i]));
                                                    // 非有限判定同高选口径
        IF aEn[i] AND (NOT _bNonFin) THEN
            IF (NOT _bFound) OR (aIn[i] < _fBest) THEN
                _fBest := aIn[i];               // 低选：严格小于才换（平值取首路）
                _uWin := INT_TO_UINT(i);        // 记胜出通道
                _bFound := TRUE;                // 已找到
            END_IF
        END_IF
    END_FOR

ELSE
    nErrId := 16#0002_03A4;         // 故障级：非法选择模式兜底
    bError := TRUE;                 // 故障码配对置位
    RETURN;                         // 直接出口（出口保持缺省无效）/ early exit

END_CASE

(* —— 段 3｜出口单点映射（名实同源） —— *)
IF _bFound THEN
    fOut := _fBest;                 // 胜出值出口
    uWin := _uWin;                  // 胜出通道出口
    bValid := TRUE;                 // 有效出口
    IF NOT _bAnyPrev THEN
        nErrId := 16#0002_0489;     // 信息级：首次有效输出沿
    END_IF
ELSE
    uWin := 0;                      // 无有效输入（哨兵零通道）
    nErrId := 16#0002_048A;         // 信息级：全通道无效
END_IF
_bAnyPrev := _bFound;               // 首次有效沿判据快照

END_FUNCTION_BLOCK

(* ---- FB_DL_ParticleCounterStat.st ---- *)
//==============================================================================
// 功能块：FB_DL_ParticleCounterStat ｜ 中文名称：尘埃粒子计数器统计与等级判定
// 所属子库：DL_Algo ｜ 版本：v1.0.0 ｜ 兼容：CODESYS V3.5+ / TwinCAT 3 / 汇川 InoProShop
// 功能描述：6 路粒径计数（0.1/0.2/0.3/0.5/1.0/5.0 微米）→ 浓度（颗每
//           立方米）→ ISO 14644-1:2015 Table 1 等级判定（生成式 Cn =
//           10^N 乘 (0.1/D)^2.08，N 允许 0.5 步进）→ 连续 N 个采样超限
//           才报警 → 失采检测。等级判定采用 Table 1 常量表锚定 + 档内
//           LOG 对数插值：** 幂运算符跨平台不可用，改用「整数档查表
//           + LOG 对数插值」，由生成式恒等式 conc/L_N = 10^(level-N)
//           保证档内插值与公式严格一致，不引入近似误差。表内「—」
//           （无限制）格跳过不参与判定。只统计与判定，不控净化设备
//           （FFU/风淋室由上位调度，本件零执行输出）。
// 开源溯源 (Origin)：道莅原创实现（参考 ISO 14644-1:2015 Table 1 公开分级口径 分类与参数域）
// 单位表：粒子计数[颗] / 采样体积[L] / 浓度[颗/m³] / 等级[—] / 采样周期[min] / 确认数[个]
// 错误码表：16#0002_3301 信息级（采样失采，等级不可判，等级清零不沿用，
//           不置 bError）/ 16#0002_3302 信息级（等级超 9 钳 9.0，或通道
//           浓度超最深有表值档且更高档无限制被表驱动跳过，不置 bError）/
//           16#0002_3305 预留禁用（不得挪用）/ 16#0002_3310 故障级（采样
//           体积小于等于 0 或组态非法，置 bError）/ 16#0002_3311 故障级
//           （浮点输入非有限，置 bError）/ 16#0002_3312 预留禁用（不得挪用）
// 状态机：E_DL_ParticleStatState（eIdle=0 / eSampling=10 / eLost=20 /
//           eFault=99），CASE 含 ELSE 兜底，ELSE 复用 3311（§3 未为本件
//           单列兜底槽，非法状态按「数据不可信」同语义处置，不得越段
//           加码）并回 eFault、等级清零（安全侧 = 不给达标假象）
// 边界行为：① 浮点输入非有限（NaN 自反判 + Inf 幅值上限判）→ 故障 3311，
//           等级清零；② fSampleVolL 小于等于防除零下限、fClassTarget 超
//           1.0~9.0 域、nConfirmSamples 超 1~10 域、tSampleTime 非正 →
//           故障 3310，先判后除防除零；③ 全通道计数为 0 且脉冲到达 =
//           合法 0 浓度，不判失采（失采只由失采定时器时间判据裁决）；
//           ④ 失采（间隔超 2 倍采样周期）→ 信息 3301 + 等级清零 +
//           bValid := FALSE，禁止沿用旧等级（旧等级会让洁净室误报达标）；
//           bOverLimit 报警锁存保持（已确认的超限事实不因失采被掩盖，
//           恢复采样后由新数据重新裁决）；⑤ 等级超 9 → 判 9.0 并信息
//           3302；⑥ 通道浓度超该通道最深有表值档且更高档为「—」→ 该
//           通道表驱动跳过不参与判定并信息 3302（披露：跳过通道的更高
//           污染贡献不参与最严等级裁决，靠 3302 可观测提示，若全通道
//           均被跳过则等级判不可用）；⑦ 上电首拍 bValid := FALSE；
//           ⑧ 失能 → eIdle、等级清零、报警清除；⑨ 失采定时器经脉冲沿
//           「断输入一拍」重启计时，失采门槛严格等于 2 倍采样周期
//           （R40 家族）。
// 修订历史：v1.0.0 2026-11-17 首版（R25 派单 · §4.2）
//==============================================================================
(*------------------------------------------------------------------------------
 * 枚举: E_DL_ParticleStatState（归属 DL_Algo，与 FB_DL_ParticleCounterStat 同文件）
 *----------------------------------------------------------------------------*)
TYPE E_DL_ParticleStatState :
(
    eIdle     := 0,    // 失能/待机：等级输出 0，报警清零 / Idle: class zeroed, alarm cleared
    eSampling := 10,   // 采样有效：最近一次脉冲已判定，等级可用 / Sampling: last pulse judged, class usable
    eLost     := 20,   // 失采：超 2 倍采样周期无脉冲，等级不可判 / Lost: no pulse within twice the sample period
    eFault    := 99    // 故障兜底态：组态非法或非有限，等级清零 / Fault fallback: config invalid or non-finite, class zeroed
);
END_TYPE
FUNCTION_BLOCK FB_DL_ParticleCounterStat
VAR_INPUT
    auCounts        : ARRAY[0..5] OF UDINT;    // 本采样周期各粒径计数 [颗]，通道序 0.1/0.2/0.3/0.5/1.0/5.0 微米 / counts per channel [particles], channels 0.1/0.2/0.3/0.5/1.0/5.0 um
    fSampleVolL     : LREAL := 1.0;            // 采样体积 [L]，域大于 0 / Sample volume [L], domain > 0
    bSamplePulse    : BOOL;                    // 采样周期完成脉冲，上升沿取数 / Sample-complete pulse, latched on rising edge
    fClassTarget    : LREAL := 7.0;            // 目标等级 [—]，1.0~9.0，0.5 步进 / Target class, 1.0~9.0, 0.5 steps
    nConfirmSamples : INT := 3;                // 连续超限确认数 [个]，1~10 / Consecutive over-limit confirmations, 1~10
    tSampleTime     : TIME := T#1M;            // 采样周期 [min]，用于失采判定 / Sample period [min], loss detection basis
    bEnable         : BOOL;                    // 总使能 / Master enable
    bReset          : BOOL;                    // 复位，上升沿清状态与计数 / Reset, rising edge clears state and counters
END_VAR
VAR_OUTPUT
    afConcM3        : ARRAY[0..5] OF LREAL;    // 各粒径浓度 [颗/m³] / Concentration per channel [particles/m3]
    fClassMeasured  : LREAL;                   // 实测等级 [—]，0.0 = 不可判 / Measured class, 0.0 = not judgeable
    bClassOk        : BOOL;                    // 实测等级不超过目标等级 / Measured class within target
    bOverLimit      : BOOL;                    // 连续确认后的超限报警锁存 / Confirmed over-limit alarm latch
    bSampleLost     : BOOL;                    // 失采标志 / Sample-loss flag
    tSinceSample    : TIME;                    // 距上次成功采样耗时 [min] / Time since last accepted sample [min]
    uSampleCount    : UDINT;                   // 累计采样次数 [次]，饱和计数 / Cumulative sample count, saturated
    uOverCount      : UDINT;                   // 累计超限报警次数 [次]，饱和计数 / Cumulative over-limit alarm count, saturated
    eErr            : UDINT;                   // 错误码，0 = 无错，码位 16#0002_3301 起信息级、16#0002_3310 起故障级（分带见错误码表） / Error code, 0 = no error, band info/fault per the code table
    bError          : BOOL;                    // 故障级标志，仅故障级错误置位 / Fault-class flag, set only on fault-level codes
    bValid          : BOOL;                    // 等级数据可用标志，失能/失采/故障闸显式 FALSE / Class data usable flag, explicit FALSE on disable/lost/fault gates
    eState          : E_DL_ParticleStatState;  // 主状态机当前状态 / Current state of the main state machine
END_VAR
VAR
    fbPulse         : R_TRIG;                  // 采样脉冲上升沿检测实例 / Sample pulse rising edge detector
    fbReset         : R_TRIG;                  // 复位上升沿检测实例 / Reset rising edge detector
    fbLostTimer     : TON;                     // 失采定时器：脉冲沿断输入一拍重启计时 / Loss timer: input broken one scan per pulse edge
    bTimerKick      : BOOL;                    // 定时器断输入一拍标志（重启计时，R40 家族）/ One-scan timer kick flag, restarts timing
    auLatch         : ARRAY[0..5] OF UDINT;    // 脉冲沿锁存的计数副本 [颗] / Latched counts copy [particles]
    fVolM3          : LREAL;                   // 采样体积换算 [m³] / Sample volume converted [m3]
    uCh             : INT;                     // 通道循环索引 [—] / Channel loop index
    nClass          : INT;                     // 等级档循环索引 [—] / Class row loop index
    fLimit          : LREAL;                   // 当前档表值 [颗/m³]，负数 = 无限制 / Table limit at current class [particles/m3], negative = no limit
    fLimitFloor     : LREAL;                   // 该通道最深有表值 [颗/m³] / Deepest limited table value of the channel
    nClassFloor     : INT;                     // 该通道最深有表值档号 [—] / Deepest limited class number of the channel
    fChLevel        : LREAL;                   // 通道判定等级 [—] / Per-channel judged class
    bAnyJudged      : BOOL;                    // 本采样是否存在参与判定的通道 / Whether any channel was judged this sample
    bClampHigh      : BOOL;                    // 本采样发生等级钳 9 或表驱动跳过 / Clamp-to-9 or table-skip occurred this sample
    nConsec         : INT;                     // 连续超限计数 [个] / Consecutive over-limit counter
END_VAR
VAR CONSTANT
    DL_PC_ZERO      : LREAL := 0.0;            // 零值常量，避免裸字面量 [—] / Zero constant, avoids a bare literal
    DL_PC_INF       : LREAL := 1.7976931348623157E308;  // LREAL 幅值上限，Inf 判据 / LREAL magnitude ceiling, Inf criterion
    DL_PC_VOL_MIN   : LREAL := 1.0E-9;         // 体积防除零下限 [L]，低于判组态非法 / Volume floor for zero-division guard [L]
    DL_PC_LITRE_M3  : LREAL := 1000.0;         // 升转立方米系数 [L/m³] / Litre-to-m3 factor
    DL_PC_CLASS_MAX : LREAL := 9.0;            // ISO 等级上限 [—] / ISO class ceiling
    DL_PC_CLASS_MIN : LREAL := 1.0;            // ISO 等级下限 [—] / ISO class floor
    DL_PC_TOL       : LREAL := 1.0E-6;         // 浮点比较容差 [—] / Float comparison tolerance
    DL_PC_CNT_MAX   : UDINT := 16#FFFF_FFFE;   // 饱和计数上限 [次] / Saturating counter ceiling
    DL_PC_LOSS_MULT : INT := 2;                // 失采判据倍率 [倍]，超 2 倍采样周期 / Loss multiplier, twice the sample period
    DL_PC_TIME_ZERO : TIME := T#0S;            // 时间零值基准 [s] / Time zero reference
END_VAR

(*------------------------------------------------------------------------------
 * ISO 14644-1:2015 Table 1 常量上限表：行 = 等级 1..9，列 = 通道
 * 0.1/0.2/0.3/0.5/1.0/5.0 微米；-1.0 = 「—」（无限制），该格跳过不参与
 * 判定。公共领域常量表，数值为标准原文（颗/m³）。
 *----------------------------------------------------------------------------*)
VAR CONSTANT
    DL_PCNT_CODE_INFO_1 : UDINT := 16#0002_3301;   // 信息级槽 1（采样失采） / info slot 1
    DL_PCNT_CODE_INFO_2 : UDINT := 16#0002_3302;   // 信息级槽 2（等级钳 9 或表驱动跳过） / info slot 2
    DL_PCNT_CODE_RSV_1  : UDINT := 16#0002_3305;   // 预留禁用（不得挪用） / reserved, do not use
    DL_PCNT_CODE_FLT_1  : UDINT := 16#0002_3310;   // 故障级槽 1（体积非正或组态非法） / fault slot 1
    DL_PCNT_CODE_FLT_2  : UDINT := 16#0002_3311;   // 故障级槽 2（输入非有限） / fault slot 2
    DL_PCNT_CODE_RSV_2  : UDINT := 16#0002_3312;   // 预留禁用（不得挪用） / reserved, do not use
    DL_PCNT_ISO_LIM : ARRAY[1..9, 0..5] OF LREAL := [
        10.0,      2.0,      -1.0,     -1.0,     -1.0,     -1.0,       // 等级 1 行 / class 1 row
        100.0,     24.0,     10.0,     4.0,      -1.0,     -1.0,       // 等级 2 行 / class 2 row
        1000.0,    237.0,    102.0,    35.0,     8.0,      -1.0,       // 等级 3 行 / class 3 row
        10000.0,   2370.0,   1020.0,   352.0,    83.0,     -1.0,       // 等级 4 行 / class 4 row
        100000.0,  23700.0,  10200.0,  3520.0,   832.0,    29.0,       // 等级 5 行 / class 5 row
        1000000.0, 237000.0, 102000.0, 35200.0,  8320.0,   293.0,      // 等级 6 行 / class 6 row
        -1.0,      2370000.0, 1020000.0, 352000.0, 83200.0, 2930.0,   // 等级 7 行，0.1 微米无限制 / class 7 row, 0.1 um unlimited
        -1.0,      23700000.0, 10200000.0, 3520000.0, 832000.0, 29300.0, // 等级 8 行，0.1 微米无限制 / class 8 row, 0.1 um unlimited
        -1.0,      -1.0,     -1.0,     35200000.0, 8320000.0, 293000.0  // 等级 9 行，0.1/0.2/0.3 微米无限制 / class 9 row, 0.1/0.2/0.3 um unlimited
    ];
END_VAR

(*------------------------------------------------------------------------------
 * 段 1｜无条件刷新区（红线 5）：三实例在任何分支之外周期调用
 *----------------------------------------------------------------------------*)
fbReset(CLK := bReset);                        // 复位沿检测无条件刷新 / reset edge refreshed unconditionally
fbPulse(CLK := bSamplePulse);                  // 采样沿检测无条件刷新 / sample edge refreshed unconditionally
bTimerKick := fbPulse.Q;                       // 本拍有脉冲则断定时器输入一拍 / break the loss timer input on pulse edge
fbLostTimer(IN := bEnable AND NOT bTimerKick,  // 断输入一拍重启计时（R40 家族）/ break input one scan to restart timing
            PT := tSampleTime * DL_PC_LOSS_MULT);  // 失采门槛 = 2 倍采样周期 / loss threshold = twice the sample period
tSinceSample := fbLostTimer.ET;                // 距上次采样耗时出口 / elapsed since last sample

(*------------------------------------------------------------------------------
 * 段 2｜复位沿：状态回 eIdle、计数清零、报警清除（改写置于沿后，防吞沿 R39）
 *----------------------------------------------------------------------------*)
IF fbReset.Q THEN
    eState      := E_DL_ParticleStatState.eIdle;
    eErr        := 16#0000_0000;               // 复位清码 / reset clears code
    bError      := FALSE;                      // 复位清故障 / reset clears fault
    fClassMeasured := DL_PC_ZERO;              // 等级清零 / class zeroed
    bClassOk    := FALSE;                      // 达标标志清除 / pass flag cleared
    bOverLimit  := FALSE;                      // 报警锁存清除 / alarm latch cleared
    bSampleLost := FALSE;                      // 失采标志清除 / loss flag cleared
    nConsec     := 0;                          // 连续超限计数清零 / consecutive counter zeroed
    uSampleCount := 0;                         // 采样计数清零 / sample count zeroed
    uOverCount  := 0;                          // 报警计数清零 / alarm count zeroed
    FOR uCh := 0 TO 5 DO
        afConcM3[uCh] := DL_PC_ZERO;           // 浓度出口清零 / concentration outputs zeroed
    END_FOR
END_IF

(*------------------------------------------------------------------------------
 * 段 3｜非有限输入闸（浮点引脚逐个：NaN 自反判 + Inf 幅值上限判，R79）
 *----------------------------------------------------------------------------*)
IF (fSampleVolL <> fSampleVolL) OR (ABS(fSampleVolL) >= DL_PC_INF)
   OR (fClassTarget <> fClassTarget) OR (ABS(fClassTarget) >= DL_PC_INF) THEN
    eState  := E_DL_ParticleStatState.eFault;
    eErr    := DL_PCNT_CODE_FLT_2;                 // 故障级：浮点输入非有限 / fault: non-finite float input
    bError  := TRUE;                           // 故障级必置 bError（R45 配对）/ fault-class pairs with bError
    bValid  := FALSE;                          // 输出不可用 / outputs unusable
    fClassMeasured := DL_PC_ZERO;              // 等级清零安全侧 / class zeroed, safe side
    bClassOk := FALSE;                         // 达标标志清除 / pass flag cleared
    bSampleLost := FALSE;                      // 故障态下失采语义让位非有限故障 / loss flag yields to non-finite fault
    RETURN;
END_IF

(*------------------------------------------------------------------------------
 * 段 4｜组态合法性闸（体积先判后除、目标域、确认数域、采样周期域）
 *----------------------------------------------------------------------------*)
IF (fSampleVolL <= DL_PC_VOL_MIN)
   OR (fClassTarget < DL_PC_CLASS_MIN - DL_PC_TOL) OR (fClassTarget > DL_PC_CLASS_MAX + DL_PC_TOL)
   OR (nConfirmSamples < 1) OR (nConfirmSamples > 10)
   OR (tSampleTime <= DL_PC_TIME_ZERO) THEN
    eState  := E_DL_ParticleStatState.eFault;
    eErr    := DL_PCNT_CODE_FLT_1;                 // 故障级：体积小于等于 0 或组态非法 / fault: volume non-positive or config invalid
    bError  := TRUE;                           // 故障级必置 bError（R45 配对）/ fault-class pairs with bError
    bValid  := FALSE;                          // 输出不可用 / outputs unusable
    fClassMeasured := DL_PC_ZERO;              // 等级清零，不给达标假象 / class zeroed
    bClassOk := FALSE;                         // 达标标志清除 / pass flag cleared
    bSampleLost := FALSE;                      // 故障态下失采语义让位组态故障 / loss flag yields to config fault
    RETURN;
END_IF

(*------------------------------------------------------------------------------
 * 段 5｜状态机：CASE 含 ELSE 兜底（非法状态 → 复用 3311 兜底 + 等级清零）
 *----------------------------------------------------------------------------*)
CASE eState OF

    E_DL_ParticleStatState.eIdle:
        fClassMeasured := DL_PC_ZERO;          // 待机等级清零 / class zeroed in idle
        bClassOk := FALSE;                     // 达标标志清除 / pass flag cleared
        bOverLimit := FALSE;                   // 报警清除 / alarm cleared
        bSampleLost := FALSE;                  // 失采标志清除 / loss flag cleared
        bValid := FALSE;                       // 失能闸显式不可用（R72）/ explicit FALSE on disable gate
        eErr := 16#0000_0000;                  // 待机无错 / no error in idle
        bError := FALSE;                       // 待机无故障 / no fault in idle
        IF bEnable THEN
            eState := E_DL_ParticleStatState.eSampling;  // 使能即进采样态，等首个脉冲 / enable enters sampling
        END_IF

    E_DL_ParticleStatState.eSampling:
        bValid := FALSE;                       // 默认不可用，脉冲判定通过才置位 / default unusable until judged
        bSampleLost := FALSE;                  // 采样态失采标志复位 / loss flag reset in sampling state
        IF fbLostTimer.Q THEN
            eState      := E_DL_ParticleStatState.eLost;   // 失采转出 / enter lost state
            bSampleLost := TRUE;               // 失采标志置位 / loss flag set
        ELSIF fbPulse.Q THEN
            uSampleCount := uSampleCount + 1;  // 采样计数递增 / increment sample count
            IF uSampleCount >= DL_PC_CNT_MAX THEN
                uSampleCount := DL_PC_CNT_MAX; // 饱和防回绕 / saturate to avoid wrap
            END_IF
            fVolM3 := fSampleVolL / DL_PC_LITRE_M3;  // 升转立方米，fSampleVolL 已闸大于 0 / litre to m3, divisor gated
            FOR uCh := 0 TO 5 DO
                auLatch[uCh]  := auCounts[uCh];                // 锁存计数副本 / latch counts
                afConcM3[uCh] := UDINT_TO_LREAL(auLatch[uCh]) / fVolM3;  // 浓度 = 计数/体积，除子已闸 / concentration, divisor gated
            END_FOR
            fClassMeasured := DL_PC_ZERO;      // 等级初始化，各通道最严（小数值优先）/ class init, strictest channel wins
            bAnyJudged     := FALSE;           // 参与判定通道存在标志复位 / any-judged flag reset
            bClampHigh     := FALSE;           // 本采样钳位/跳过标志复位 / clamp-or-skip flag reset
            FOR uCh := 0 TO 5 DO
                nClassFloor := 0;              // 最深有表值档复位 / deepest limited class reset
                fLimitFloor := DL_PC_ZERO;     // 最深有表值复位 / deepest limited value reset
                FOR nClass := 1 TO 9 DO
                    fLimit := DL_PCNT_ISO_LIM[nClass, uCh];  // 查表取当前档上限 / table lookup
                    IF fLimit >= DL_PC_ZERO THEN
                        nClassFloor := nClass; // 记录最深有表值档 / track deepest limited class
                        fLimitFloor := fLimit; // 记录最深有表值 / track deepest limited value
                    END_IF
                END_FOR
                IF afConcM3[uCh] > fLimitFloor THEN
                    bClampHigh := TRUE;        // 超最深有表值档 → 表驱动跳过或钳 9 / beyond deepest limited row
                    IF nClassFloor >= 9 THEN
                        IF fClassMeasured < DL_PC_CLASS_MAX THEN
                            fClassMeasured := DL_PC_CLASS_MAX;  // 等级超 9 → 钳 9.0 / beyond class 9, clamp
                        END_IF
                        bAnyJudged := TRUE;    // 钳 9 视为参与判定 / clamp counts as judged
                    END_IF
                    // 更高档无表值（nClassFloor < 9）→ 本通道跳过不参与判定，仅提示（边界行为⑥）
                ELSIF afConcM3[uCh] > DL_PC_TOL THEN
                    fChLevel := LREAL(nClassFloor) + LOG(afConcM3[uCh] / fLimitFloor);  // 档内/档下对数插值，生成式恒等口径 / in-row log interpolation, exact per the generation formula
                    IF fChLevel > fClassMeasured THEN
                        fClassMeasured := fChLevel;  // 取最严（小数值等级更严）/ strictest (smallest number) wins
                    END_IF
                    bAnyJudged := TRUE;        // 存在参与判定通道 / a channel was judged
                END_IF
                // 浓度为 0 → 合法零浓度，等级 0，不参与拉高最严值 / zero concentration is legal
            END_FOR
            bClassOk := bAnyJudged AND (fClassMeasured <= fClassTarget + DL_PC_TOL);  // 达标判定（容差比较，禁浮点判等），全通道跳过时不可判 / pass judgement with tolerance, not judgeable when all channels skipped
            IF NOT bAnyJudged THEN
                bClassOk := FALSE;             // 全通道跳过 → 等级不可判 / all channels skipped, class not judgeable
                bValid := FALSE;               // 输出不可用 / outputs unusable
            ELSE
                bValid := TRUE;                // 等级数据可用 / class data usable
            END_IF
            IF bClassOk THEN
                nConsec := 0;                  // 达标清连续计数 / pass resets consecutive counter
            ELSE
                nConsec := nConsec + 1;        // 超限连续计数递增 / over-limit increments counter
                IF nConsec >= nConfirmSamples THEN
                    IF NOT bOverLimit THEN
                        uOverCount := uOverCount + 1;  // 新报警事件计数 / new alarm event counted
                        IF uOverCount >= DL_PC_CNT_MAX THEN
                            uOverCount := DL_PC_CNT_MAX;  // 饱和防回绕 / saturate to avoid wrap
                        END_IF
                    END_IF
                    bOverLimit := TRUE;        // 连续确认后置报警锁存 / alarm latch after confirmation
                END_IF
            END_IF
            eErr   := 16#0000_0000;            // 采样有效，先清码 / valid sample clears code first
            IF bClampHigh THEN
                eErr := DL_PCNT_CODE_INFO_2;   // 信息级：等级钳 9 或表驱动跳过 / info: clamped or table-skipped
            END_IF
            bError := FALSE;                   // 信息级不置 bError / info never raises bError
        END_IF

    E_DL_ParticleStatState.eLost:
        bValid := FALSE;                       // 失采闸显式不可用（R72）/ explicit FALSE on lost gate
        fClassMeasured := DL_PC_ZERO;          // 禁止沿用旧等级，等级清零 / never keep old class, zeroed
        bClassOk := FALSE;                     // 达标标志清除 / pass flag cleared
        eErr   := DL_PCNT_CODE_INFO_1;             // 信息级：采样失采 / info: sample lost
        bError := FALSE;                       // 信息级不置 bError / info never raises bError
        bSampleLost := TRUE;                   // 失采态期间标志保持 / loss flag held in lost state
        IF fbPulse.Q THEN
            eState := E_DL_ParticleStatState.eSampling;  // 事件沿退出 / exit on pulse edge
            bSampleLost := FALSE;              // 前置（失采定时器 Q）随断输入一拍消失 / precondition clears with the timer kick
            eErr := 16#0000_0000;              // 恢复清码 / clear code on recovery
        END_IF

    ELSE
        eState := E_DL_ParticleStatState.eFault;  // 非法状态兜底 / illegal-state fallback
        eErr   := DL_PCNT_CODE_FLT_2;              // 兜底复用故障级槽 2（数据不可信同语义，§3 未单列兜底槽，不得越段加码）/ fallback reuses fault slot 2, no out-of-band code
        bError := TRUE;                        // 故障级必置 bError / fault-class pairs with bError
        bValid := FALSE;                       // 输出不可用 / outputs unusable
        fClassMeasured := DL_PC_ZERO;          // 等级清零安全侧 / class zeroed, safe side
        bClassOk := FALSE;                     // 达标标志清除 / pass flag cleared
END_CASE
END_FUNCTION_BLOCK

(* ---- FB_DL_PeakHoldFilter.st ---- *)
(*==============================================================================
 * 组件名称 (Component)  : FB_DL_PeakHoldFilter
 * 所属子库 (Sublibrary) : DL_Algo
 * 当前版本 (Version)    : 1.0.0
 * 兼容性   (Platform)   : CODESYS 3.5+ / TwinCAT 3 / 汇川 InoProShop / 施耐德 Machine Expert
 *                         仅依赖 Standard.library（TON / TIME_TO_REAL），零厂商私有库
 * 功能描述 (Function)   : 峰值保持（peak hold）。持续跟踪输入最大值；保持时长 tHoldTime
 *                         内无新的更高峰值即自动回落（回落到当前输入值），随后转为跟随输入。
 *                         典型用途：液压冲击峰值记录、张力瞬时峰值捕获、压力尖峰监测。
 *                         保持计时用 TON 事件重启式：每当新峰值出现，本拍把 TON 的 IN
 *                         强制为 FALSE 一拍，TON 内部 ET/Q 即复位（比外部清零更稳，
 *                         不依赖调用方沿信号）；其余拍 IN = bHolding。
 * 接口     (Interface)  : 输入 bEnable 使能、bReset 复位峰值、fIn 采样输入 [EU]、
 *                         tHoldTime 峰值保持时长 [s]；
 *                         输出 fPeak 保持峰值 [EU]、bHolding 是否处于保持期、
 *                         tHoldElapsed 已保持时长 [s]、bValid 输出有效、bError、uErrorId。
 * 边界     (Boundary)   : ① 属主边界：只做峰值保持，不做峰值-时间戳归档（另件）。
 *                         ② 非有限输入 → 进故障态冻结输出，uErrorId=16#0004_0002；
 *                         恢复路径：bEnable=FALSE 或 bReset=TRUE。
 *                         ③ tHoldTime < 0 判参数非法（TIME 无负值语义，钳到 T#0S 并置信息码
 *                         16#0004_0001）；tHoldTime = T#0S 表示不保持，逐拍跟随输入。
 *                         ④ **TON 无条件每周期调用**（R7）：位于 CASE 之外的段 3，
 *                         与状态机解耦，任何状态下计时器都被刷新。
 *                         ⑤ 零全局耦合（无 GVL / VAR_EXTERNAL / 物理地址）。
 * 分工声明 (Scope)      : 与 `FB_DL_HoldLastGoodFilter` 分工：坏值保持归那件、
 *                         峰值保持归本件；与 `FB_DL_RateOfChangeFilter` 分工：斜率限幅归那件。
 * 来源标签 (Source Tag) : 原创实现（无外部代码引入）
 * 码表     (Codes)      : 16#0004_0000 无故障 / 16#0004_0001 保持时长非法已钳位（信息级）/
 *                         16#0004_0002 输入非有限（故障级）/ 16#0004_0005 非法状态（故障级）。
 * 红线自检 (Redline)    : R1 ✓ 零 GVL/VAR_EXTERNAL ｜ R2 ✓ 零 %I/%Q/%M ｜ R3 ✓ 纯 IEC 61131-3
 *                         R4 ✓ 非有限拒绝 + 时长域闸 + 无除法 ｜ R5 ✓ 声明逐行同行双语注释
 *                         R6 ✓ 四态 ENUM + CASE + ELSE 兜底 ｜ R7 ✓ TON 实例 CASE 外无条件刷新
 * 修订历史 (Revision)   : 2026-11-23  v1.0.0  R77 首版（批次 B3 · 序号 10）
 * 验收向量 (Acceptance) : ① tHoldTime=T#1S，输入 5.0 后降到 3.0 → fPeak 保持 5.0，
 *                         bHolding=TRUE；保持期满后 fPeak 回落到 3.0；
 *                         ② bReset=TRUE 一拍 → fPeak 立即等于当前 fIn，bHolding=TRUE；
 *                         ③ tHoldTime=T#0S → 逐拍跟随输入，fPeak = fIn（不保持）；
 *                         ④ fIn=Inf → uErrorId=16#0004_0002，bError=TRUE，fPeak 冻结；
 *                         ⑤ bEnable=FALSE → fPeak 冻结，bValid=FALSE，计时器照常刷新。
 *==============================================================================*)

(*-----------------------------------------------------------------------------
 * 枚举: E_DL_PeakHoldState（峰值保持状态机，归属 DL_Algo，与本件同文件，全库唯一属主）
 *----------------------------------------------------------------------------*)
TYPE E_DL_PeakHoldState :
(
    eInit  := 0,    // 首扫 / 复位后：峰值取当前输入 / First scan or after reset: peak equals input
    eRun   := 10,   // 运行态：捕获更高峰并重启保持计时 / Running: capture higher peaks and restart timer
    eHold  := 20,   // 保持态：未使能，输出冻结 / Hold: disabled, output frozen
    eFault := 99    // 故障态：输出冻结，等待 bEnable 跌落或 bReset / Fault: frozen until cleared
);
END_TYPE

FUNCTION_BLOCK FB_DL_PeakHoldFilter
VAR_INPUT
    bEnable   : BOOL := FALSE;      // 使能，FALSE 冻结峰值 / Enable, FALSE freezes the peak
    bReset    : BOOL := FALSE;      // 复位峰值到当前输入（单拍有效） / Reset peak to current input, single scan
    fIn       : LREAL := 0.0;       // 采样输入 [EU] / Sampling input [EU]
    tHoldTime : TIME := T#1S;       // 峰值保持时长，T#0S = 不保持 [s] / Peak hold duration, zero means follow
END_VAR
VAR_OUTPUT
    fPeak        : LREAL;   // 保持峰值 [EU] / Held peak [EU]
    bHolding     : BOOL;    // 是否处于保持期 [-] / Whether inside the hold window
    tHoldElapsed : TIME;    // 已保持时长 [s] / Elapsed hold duration
    bValid       : BOOL;    // 输出有效标志 [-] / Output valid flag
    bError       : BOOL;    // 故障标志，与 uErrorId 联动 [-] / Fault flag coupled with uErrorId
    uErrorId     : UDINT;   // 故障码，0 = 无故障 [-] / Error code, zero means healthy
END_VAR
VAR
    tonHold  : TON;                 // 峰值保持计时器（无条件每周期刷新） / Peak hold timer, refreshed unconditionally
    _bRstPul : BOOL;                // 新峰值事件脉冲（本拍重启计时） [-] / New-peak event pulse for timer restart
    _bNewPk  : BOOL;                // 本拍出现更高峰 [-] / Higher peak appeared this scan
    eState   : E_DL_PeakHoldState;  // 状态机当前状态 [-] / Current state
END_VAR
VAR CONSTANT
    DL_PHF_ZERO_L : LREAL := 0.0;   // 零基准（含非有限判零） [-] / Zero base including non-finite probe
    DL_PHF_ZERO_T : TIME := T#0S;   // 时长零基准 [s] / Zero duration base
END_VAR

(* —— 段 1：参数域闸（时长非负；TIME 无负值，仍显式判等以防方言差异） —— *)
uErrorId := 16#0004_0000;                          // 预置无故障 / Preset healthy
IF tHoldTime < DL_PHF_ZERO_T THEN
    tHoldTime := DL_PHF_ZERO_T;                    // 负时长钳到零 / Negative duration clamped to zero
    uErrorId  := 16#0004_0001;                     // 信息级：保持时长已钳位 / Info: hold duration clamped
END_IF

(* —— 段 2：非有限输入防御（进故障态冻结输出） —— *)
IF (fIn <> fIn) OR ((fIn - fIn) <> DL_PHF_ZERO_L) THEN
    eState   := eFault;                            // 强制故障态 / Force fault state
    uErrorId := 16#0004_0002;                      // 故障级：输入非有限 / Fault: non-finite input
END_IF

(* —— 段 3：新峰值检测与计时器重启脉冲（仅在使能且运行态有效） —— *)
_bNewPk  := FALSE;                                 // 每拍清零事件位 / Clear event flag every scan
_bRstPul := FALSE;
IF bEnable AND (eState <> eFault) THEN
    IF fIn > fPeak THEN
        _bNewPk  := TRUE;                          // 出现更高峰 / Higher peak detected
        _bRstPul := TRUE;                          // 本拍强制 TON 的 IN=FALSE 以复位 ET/Q / Force timer reset
    END_IF
END_IF

(* —— 段 4：复位请求 → 回首扫（峰值对齐当前输入） —— *)
IF bReset THEN
    eState := eInit;
END_IF

(* —— 段 5：状态派生 —— *)
IF NOT bEnable THEN
    eState := eHold;                               // 未使能：冻结 / Disabled: freeze
ELSIF eState = eFault THEN
    eState := eFault;                              // 故障态保持 / Fault holds
ELSIF eState = eInit THEN
    eState := eInit;                               // 首扫保持一拍 / Init holds one scan
ELSE
    eState := eRun;
END_IF

(* —— 段 6：计时器无条件每周期刷新（R7 硬要求，位于 CASE 之外） —— *)
(* IN 在「使能 且 处于保持中 且 本拍无新峰」时为 TRUE；新峰拍强制 FALSE 完成复位 *)
(* IN is TRUE only when enabled, holding, and no new peak this scan; a new peak forces FALSE to reset *)
tonHold(IN := bEnable AND (eState <> eFault) AND (NOT _bRstPul), PT := tHoldTime);

(* —— 段 7：主状态机（CASE 覆盖 + ELSE 兜底） —— *)
CASE eState OF

    eInit:
        fPeak        := fIn;                       // 峰值对齐当前输入 / Align peak with input
        bHolding     := TRUE;                      // 进入保持期 / Enter hold window
        tHoldElapsed := tonHold.ET;
        bValid       := TRUE;
        eState       := eRun;

    eRun:
        IF _bNewPk THEN
            fPeak := fIn;                          // 捕获更高峰 / Capture higher peak
        ELSIF tonHold.Q THEN
            fPeak := fIn;                          // 保持期满：回落到当前输入 / Hold expired: fall back to input
        END_IF
        bHolding     := NOT tonHold.Q;             // 期满后不再处于保持期 / No longer holding after expiry
        tHoldElapsed := tonHold.ET;
        bValid       := TRUE;

    eHold:
        (* 未使能：峰值与计时保持冻结，恢复使能后继续 / Disabled: peak and timer frozen *)
        tHoldElapsed := tonHold.ET;
        bValid       := FALSE;

    eFault:
        (* 故障态：峰值冻结（不推 0，避免下游误判），计时器仍刷新 / Fault: peak frozen, timer still refreshed *)
        tHoldElapsed := tonHold.ET;
        bValid       := FALSE;

    ELSE
        eState   := eFault;
        bValid   := FALSE;
        uErrorId := 16#0004_0005;                  // 故障级：非法状态 / Fault: illegal state

END_CASE;

(* —— 段 8：出口映射（bError 与 uErrorId 同源；信息级 16#0004_0001 不置 bError） —— *)
bError := (uErrorId <> 16#0004_0000) AND (uErrorId <> 16#0004_0001);

END_FUNCTION_BLOCK

(* ---- FB_DL_PeltierTempCtrl.st ---- *)
(*
  道莅工业代码库 | DL_Algo | FB_DL_PeltierTempCtrl
  版本: 1.0.0 | 日期: 2026-11-23 | 轮次: R75
  开源溯源: self-cleanroom（无外部来源；行业池·精密温控 TEC 语义，零代码行复制）
  功能: 半导体制冷（TEC）双向温控——单 PI 输出带符号（正=加热极性/负=制冷极性），
        极性切换带回差（fDeadband）与最短驻留（tPolDwell，经 eSwitch 过渡相强制
        输出归零泄流），双向抗饱和（限幅同向禁积分）。
  兼容性: CODESYS 3.5 / TwinCAT 3 / 汇川 InoProShop；仅依赖标准 TON / R_TRIG / LIMIT，零厂商私有库
  接口: 输入使能/温度设定/实测/PI 增益/输出限幅/积分限幅/切换回差/极性驻留/
        周期/复位；输出 fOutPct [%，-100..100]/bHeatMode/bCoolMode/fErrC/
        eState/eCause/bError/nErrId。
  码表: 16#0002_030B 故障级：温控故障总码（组态非法/温度非有限，锁存至复位沿）
        16#0002_0400 信息级：极性切换过渡进入（eSwitch 相，输出强制归零泄流）
        码段说明：0002 段故障子带 03xx / 信息子带 04xx，槽位经全库实扫空闲。
  边界: ① 极性切换三闸：误差越反向回差 ∧ 极性驻留满 tPolDwell ∧ 使能保持；
        切换经 eSwitch 过渡相（输出归零一拍周期 tPolDwell 泄流）后按当拍误差
        符号落极；
        ② 抗饱和：输出已饱和且误差继续同向 → 本拍不积分（双向对称口径）；
        ③ 极性驻留计时 tonDwell IN 挂加热/制冷相，经 eSwitch（IN 假）自然复位
        （R188 自复位口径）；
        ④ 温度/设定 NaN 故障锁存，输出钳零（安全侧）；
        ⑤ TON/R_TRIG 段 0 无条件周期刷新；⑥ 故障解除唯一路径 = 复位沿 ∧ 组态合法；
        ⑦ 零全局耦合。
  邻件比对: PidController（通用 PID vs 本件冷热极性切换+双向抗饱和 TEC 专用件）。
  修订历史: 2026-11-23 v1.0.0 R75 首版（复杂件批 B3 · C13）
*)

TYPE E_DL_PtcState :
(
    eIdle   := 0,   // 待机（输出零） | Idle, output zero
    eHeat   := 10,  // 加热极性（输出 >= 0） | Heat polarity, output non-negative
    eCool   := 20,  // 制冷极性（输出 <= 0） | Cool polarity, output non-positive
    eSwitch := 30,  // 极性切换过渡（输出归零泄流） | Polarity switch transition, output zero
    eFault  := 90   // 故障锁存相 | Fault latch phase
);
END_TYPE

TYPE E_DL_PtcCause :
(
    eNone          := 0,  // 无故障 | No cause
    eCfgIllegal    := 1,  // 组态非法 | Illegal configuration
    eSensNonFinite := 2   // 温度信号非有限 | Temperature signal non-finite
);
END_TYPE

FUNCTION_BLOCK FB_DL_PeltierTempCtrl
VAR_INPUT
    bEn        : BOOL := FALSE;    // 温控使能 [-] | Control enable
    fTempSp    : REAL := 25.0;     // 温度设定 [°C] | Temperature setpoint
    fTempAct   : REAL := 25.0;     // 温度实测 [°C] | Temperature actual
    fKp        : REAL := 20.0;     // 比例增益，域 > 0 [%/°C] | Proportional gain
    fKi        : REAL := 4.0;      // 积分增益，域 >= 0 [%/(°C·s)] | Integral gain
    fOutMax    : REAL := 100.0;    // 输出限幅，域 > 0 [%] | Output limit
    fIntLim    : REAL := 50.0;     // 积分限幅，域 (0, fOutMax] [%] | Integral limit
    fDeadband  : REAL := 0.5;      // 极性切换回差，域 >= 0 [°C] | Polarity switch hysteresis
    tPolDwell  : TIME := T#2S;     // 极性最短驻留/过渡泄流时长，域 > T#0S | Polarity dwell and transition time
    fDtSec     : REAL := 0.1;      // 控制周期，域 (0, 1] [s] | Control cycle time
    bReset     : BOOL := FALSE;    // 复位命令，上升沿清故障 [-] | Reset command, rising edge
END_VAR
VAR_OUTPUT
    fOutPct   : REAL;               // 输出出口（带符号：正=加热/负=制冷）[%] | Signed output outlet, positive heat
    bHeatMode : BOOL;               // 加热极性态 [-] | Heat polarity state
    bCoolMode : BOOL;               // 制冷极性态 [-] | Cool polarity state
    fErrC     : REAL;               // 温差出口（Sp - Act）[°C] | Error outlet
    eState    : E_DL_PtcState;      // 状态出口 | State outlet
    eCause    : E_DL_PtcCause;      // 故障成因出口 | Fault cause outlet
    bError    : BOOL;               // 故障锁存标志 [-] | Fault latch flag
    nErrId    : UDINT;              // 事件码，0 = 无事件 | Event code, 0 = none
END_VAR
VAR
    _eState  : E_DL_PtcState := E_DL_PtcState.eIdle;   // 内部状态（CASE 唯一写入目标） | Internal state
    _eCause  : E_DL_PtcCause := E_DL_PtcCause.eNone;   // 成因锁存 | Latched cause
    _bFault  : BOOL;            // 故障锁存位 | Fault latch bit
    _fInt    : REAL := 0.0;     // 积分项内部镜像 [%] | Integral term mirror
    _fOutPct : REAL := 0.0;     // 输出内部镜像 [%] | Output mirror
    _bCfgBad : BOOL;            // 组态非法当拍量 [-] | Illegal configuration
    _bSensBad: BOOL;            // 温度信号非有限当拍量 [-] | Temperature non-finite this scan
    _uInfo   : UDINT;           // 信息码每拍重算 | Info code per scan
    fErr     : REAL;            // 温差当拍量 [°C] | Error this scan
    fRaw     : REAL;            // 未限幅输出当拍量 [%] | Raw output this scan
    rtReset  : R_TRIG;          // 复位沿实例，段 0 无条件刷新 | Reset edge instance
    tonDwell : TON;             // 极性驻留计时，段 0 无条件刷新 | Polarity dwell timer
    tonSw    : TON;             // 过渡泄流计时，段 0 无条件刷新 | Transition discharge timer
END_VAR

(* —— 段 0：当拍量派生 + 定时器与沿实例无条件周期刷新（R7 红线） —— *)
_bSensBad := (fTempSp <> fTempSp) OR (fTempAct <> fTempAct);                // 温度信号 NaN 自反判 / Temperature NaN self-reflex check
_bCfgBad := (fKp <= 0.0) OR (fKi < 0.0) OR (fOutMax <= 0.0) OR (fIntLim <= 0.0)
         OR (fIntLim > fOutMax) OR (fDeadband < 0.0) OR (tPolDwell <= T#0S)
         OR (fDtSec <= 0.0) OR (fDtSec > 1.0);                              // 组态域闸 / Configuration gate
rtReset(CLK := bReset);                                                     // 复位沿每拍必调 / Reset edge every scan
tonDwell(IN := (_eState = E_DL_PtcState.eHeat) OR (_eState = E_DL_PtcState.eCool), PT := tPolDwell); // 驻留计时挂极性相 / Dwell timer in polarity states
tonSw(IN := (_eState = E_DL_PtcState.eSwitch), PT := tPolDwell);            // 泄流计时挂过渡相 / Discharge timer in transition

(* —— 段 1：单拍量预清零 + 温差派生（待机相极性判据依赖，全相可用） —— *)
_uInfo := 16#0000_0000;                                                     // 信息码每拍重算 / Info recomputed per scan
fErr := 0.0;                                                                // 温差预清（NaN 时保持零，安全侧）/ Error preset
fRaw := 0.0;                                                                // 原始输出预清 / Raw output preset
IF (NOT _bSensBad) AND (NOT _bFault) THEN
    fErr := fTempSp - fTempAct;                                             // 温差（正=欠温需加热）[°C]，全相派生 / Error derived in all states
END_IF

(* —— 段 2：复位沿 + 组态/传感器域闸 —— *)
IF rtReset.Q AND (NOT _bCfgBad) THEN                                        // 复位沿且组态合法 / Reset with legal config
    _bFault := FALSE;                                                       // 清故障锁存位 / Clear fault latch
    _eCause := E_DL_PtcCause.eNone;                                         // 清成因 / Clear cause
    _fInt := 0.0;                                                           // 清积分（复位后重新起控） / Clear integral on reset
    IF _eState = E_DL_PtcState.eFault THEN
        _eState := E_DL_PtcState.eIdle;                                     // 故障相迁出唯一路径 / Sole fault exit
    END_IF
END_IF
IF _bCfgBad THEN                                                            // 组态域闸 / Configuration gate
    _bFault := TRUE;
    _eCause := E_DL_PtcCause.eCfgIllegal;                                   // 归因组态 / Cause: config
END_IF
IF _bSensBad AND (NOT _bFault) THEN                                         // 传感器域闸（组态闸优先归因） / Sensor gate
    _bFault := TRUE;
    _eCause := E_DL_PtcCause.eSensNonFinite;                                // 归因传感器 / Cause: sensor
END_IF

(* —— 段 3：PI 计算（双向抗饱和：限幅同向禁积分，边界②） —— *)
IF (NOT _bFault) AND bEn
   AND ((_eState = E_DL_PtcState.eHeat) OR (_eState = E_DL_PtcState.eCool)) THEN
    fRaw := fKp * fErr + _fInt;                                             // 未限幅输出 [%]（fErr 已段 1 全相派生）/ Raw output
    IF (fRaw >= fOutMax) AND (fErr > 0.0) THEN
        ;                                                                   // 加热向饱和且误差仍正向：本拍不积分 / Saturated toward heat, skip integration
    ELSIF (fRaw <= -fOutMax) AND (fErr < 0.0) THEN
        ;                                                                   // 制冷向饱和且误差仍负向：本拍不积分 / Saturated toward cool, skip integration
    ELSE
        _fInt := _fInt + fKi * fErr * fDtSec;                               // 积分递推 [%.s] / Integration step
        _fInt := LIMIT(-fIntLim, _fInt, fIntLim);                           // 积分限幅 / Integral clamp
    END_IF
    _fOutPct := LIMIT(-fOutMax, fKp * fErr + _fInt, fOutMax);               // 输出限幅 [%] / Output clamp
END_IF

(* —— 段 4：状态机（ENUM + CASE，ELSE 兜底） —— *)
CASE _eState OF

E_DL_PtcState.eIdle:
    _fOutPct := 0.0;                                                        // 待机输出零 / Idle output zero
    IF bEn AND (NOT _bFault) THEN
        IF fErr >= 0.0 THEN                                                 // 首次进入按温差符号落极（NaN 已被域闸拦） / Initial polarity by error sign
            _eState := E_DL_PtcState.eHeat;                                 // 欠温进加热极性 / Under-temperature, heat
        ELSE
            _eState := E_DL_PtcState.eCool;                                 // 过温进制冷极性 / Over-temperature, cool
        END_IF
    END_IF

E_DL_PtcState.eHeat:
    IF (NOT bEn) OR _bFault THEN
        _eState := E_DL_PtcState.eIdle;                                     // 使能撤/故障回待机 / Disable or fault, idle
    ELSIF (fErr < -fDeadband) AND tonDwell.Q THEN                           // 切换三闸：越反向回差 ∧ 驻留满 ∧ 使能（边界①）/ Three switch gates
        _uInfo := 16#0002_0400;                                             // 信息级：极性切换过渡进入 / Info: transition entered
        _eState := E_DL_PtcState.eSwitch;                                   // 进过渡相泄流 / Enter transition
    END_IF

E_DL_PtcState.eCool:
    IF (NOT bEn) OR _bFault THEN
        _eState := E_DL_PtcState.eIdle;                                     // 使能撤/故障回待机 / Disable or fault, idle
    ELSIF (fErr > fDeadband) AND tonDwell.Q THEN                            // 切换三闸（对称口径）/ Three switch gates, symmetric
        _uInfo := 16#0002_0400;                                             // 信息级：极性切换过渡进入 / Info: transition entered
        _eState := E_DL_PtcState.eSwitch;                                   // 进过渡相泄流 / Enter transition
    END_IF

E_DL_PtcState.eSwitch:
    _fOutPct := 0.0;                                                        // 过渡相输出强制归零（泄流）/ Transition output forced zero
    _fInt := 0.0;                                                           // 极性翻转清积分（防反向饱和滞后）/ Clear integral on polarity transition
    IF (NOT bEn) OR _bFault THEN
        _eState := E_DL_PtcState.eIdle;                                     // 使能撤/故障回待机 / Disable or fault, idle
    ELSIF tonSw.Q THEN
        IF fErr < 0.0 THEN
            _eState := E_DL_PtcState.eCool;                                 // 泄流毕按当拍误差落制冷极 / Discharge done, cool polarity
        ELSE
            _eState := E_DL_PtcState.eHeat;                                 // 泄流毕按当拍误差落加热极 / Discharge done, heat polarity
        END_IF
    END_IF

E_DL_PtcState.eFault:
    _fOutPct := 0.0;                                                        // 故障相输出钳零（安全侧）/ Fault output zero
    ;                                                                       // 仅段 2 复位沿可迁出 / Only reset edge leaves

ELSE
    _bFault := TRUE;                                                        // 非法状态兜底（R6）/ Illegal state fallback
    _eCause := E_DL_PtcCause.eCfgIllegal;                                   // 归因归并组态 / Cause folded to config
    _eState := E_DL_PtcState.eFault;

END_CASE

(* —— 段 5：故障锁存状态迁移闸 —— *)
IF _bFault AND (_eState <> E_DL_PtcState.eFault) THEN
    _eState := E_DL_PtcState.eFault;                                        // 锁存即入故障相 / Latch enters fault phase
END_IF

(* —— 段 6：出口单点映射（名实同源；锁存码回放） —— *)
fOutPct := _fOutPct;                                                        // 输出出口 [%] / Output outlet
bHeatMode := (_eState = E_DL_PtcState.eHeat);                               // 加热极性镜像 / Heat mirror
bCoolMode := (_eState = E_DL_PtcState.eCool);                               // 制冷极性镜像 / Cool mirror
fErrC := fErr;                                                              // 温差出口 [°C] / Error outlet
eState := _eState;                                                          // 状态出口 / State outlet
eCause := _eCause;                                                          // 成因出口 / Cause outlet
bError := _bFault;                                                          // 故障标志同源 / Error flag from latch
IF _bFault THEN
    nErrId := 16#0002_030B;                                                 // 故障锁存码回放 / Replay latched fault code
ELSE
    nErrId := _uInfo;                                                       // 信息码 / Info code
END_IF

END_FUNCTION_BLOCK

(* ---- FB_DL_PeriodicDisturbComp.st ---- *)
(*
  ==================================================================
  组件名 Component  : FB_DL_PeriodicDisturbComp
  分类   Category   : DL_Algo
  复杂度 Complexity  : cx5
  版本   Version    : 1.0.1
  功能   Purpose    : 周期性扰动重复控制补偿器。内模原理：环形延迟线按周期
                      拍数存储上周期同相位误差，泄漏积分（遗忘因子）逐拍正
                      反馈累加，收敛增益钳位后取负作为前馈补偿输出。适用轧
                      辊偏心 / 卷筒周期张力等固定周期扰动。与 DisturbanceObserver
                      非周期观测分工互引。
  来源   Source     : self（控制理论公开：重复控制 / 内模原理）
  溯源   Origin     : IEC 61131-3 标准语义的道莅防御性实现；重复控制内模为
                      公开控制理论语义，clean-room 自研实现，未复制任何厂商
                      私有库源码。
  平台   Platform   : 纯 IEC 61131-3，CODESYS / TwinCAT / InoProShop 通用
  分工声明 Split     : 与 FB_DL_DisturbanceObserver 分工——后者做非周期扰动
                      状态观测，本件做固定周期扰动的内模累积补偿；本件只
                      输出补偿量，不做误差观测器极点配置。
  作者   Author     : 道莅代码库 · PLC 编程专家（R58）
  ------------------------------------------------------------------
  边界 Boundary     :
                      一 组态域：nPeriodTicks ∈ [2..4096]（拍），fForget ∈
                         [0..0.999]（无量纲，取 1.0 会无界累积故禁用），
                         fGain ∈ [0..1.0]（无量纲）；越域锁存（解除 = bReset
                         沿，R188），锁存与失能期补偿输出安全侧零；
                      二 每次调用 = 一拍：先读后写（读上周期同相位存量，
                         写本拍泄漏积分），拍推进仅在使能且域内；
                      三 非有限误差拒收（自反双判据）：本拍环不写入、输出
                         冻结保持，拒收计数出口 nSkipCnt 供调用方可观测；
                      四 环容量固定 4096，周期组态改变时写指针按新周期回
                         绕（MOD 式比较回绕，无移位无溢出）；
                      五 无全局变量、无外部变量声明、无物理地址寻址；
                      六 维护纪律（R59 轻①）：环块双清须同步维护——凡清环块
                         _aRing 必须同时清写指针 _uWidx，首扫段与复位段两处
                         双清块增删必须同步对齐，禁止只清其一。
  修订记录 Revision  :
    2026-11-21  v1.0.0  R58 首版（批 3 · 序号 10）
    2026-11-21  v1.0.1  R59 返修轻①②：头注释补环块双清同步维护纪律（边界六）；常量 DL_PDC_SKIPMAX 名实不符
                        改名 DL_PDC_CNTMAX（计数防回绕上界，覆盖 _nTick 与 nSkipCnt 两处钳定用法）
  ==================================================================
*)

FUNCTION_BLOCK FB_DL_PeriodicDisturbComp
VAR_INPUT
    fErr        : LREAL := 0.0;   // 误差反馈输入 [工程单位] / the error feedback input [engineering unit]
    nPeriodTicks: UINT  := 100;   // 扰动周期拍数 [拍]，域 2..4096 / the disturbance period in ticks, two through four thousand ninety six
    fForget     : LREAL := 0.95;  // 遗忘因子 [无量纲]，域 0..0.999 / the forgetting factor, zero through point nine nine nine
    fGain       : LREAL := 0.5;   // 收敛增益 [无量纲]，域 0..1.0 / the convergence gain, zero through one
    bEnable     : BOOL  := FALSE; // 使能，失能输出安全侧零且环冻结 [-] / enable, disabling zeroes the output and freezes the ring
    bReset      : BOOL  := FALSE; // 复位上升沿清环与锁存 [-] / reset rising edge clears the ring and the latch
END_VAR
VAR_OUTPUT
    fComp   : LREAL := 0.0; // 补偿输出（前馈，取负反馈）[工程单位] / the compensation outlet, the negative feedforward [engineering unit]
    bLearned: BOOL := FALSE; // 环已填满一周期指示 [-] / the ring filled one period indicator
    nSkipCnt: UDINT := 0;   // 非有限拒收拍计数 [拍] / the skipped non finite tick count
    bError  : BOOL := FALSE; // 域闸故障锁存标志 [-] / the domain gate fault latch flag
END_VAR
VAR
    rtReset : R_TRIG; // 复位沿检测，段 0 无条件刷新 / the reset edge
    _aRing  : ARRAY[0..4095] OF LREAL; // 环形延迟线 [工程单位] / the ring delay line [engineering unit]
    _uWidx  : UINT := 0;   // 环写指针 [槽] / the ring write index [slot]
    _nTick  : UDINT := 0;  // 使能以来累计拍数 [拍]（填满判定）/ the ticks since enabled [tick]
    _bLatch : BOOL := FALSE; // 域闸锁存位 [-] / the domain gate latch bit
    _bInit  : BOOL := FALSE; // 首扫初始化完成标志（R310）/ the first scan flag
    _nPer   : DINT;        // 周期拍数 DINT 工作副本 [拍] / the period as a DINT work copy [tick]
    _bFin   : BOOL;        // 误差有限工作量 [-] / the error finiteness work flag
    _nI     : DINT;        // 清环遍历索引 [槽] / the ring clear loop index
END_VAR
VAR CONSTANT
    DL_PDC_PERMAX : UINT := 4096;  // 周期拍数上界 [拍]，与环容量一致 / the period bound, aligned with the ring capacity
    DL_PDC_FGTMAX : LREAL := 0.999; // 遗忘因子上界 [无量纲] / the forgetting ceiling
    DL_PDC_CNTMAX : UDINT := 4294967294; // 计数防回绕上界 [拍]（R59 轻②：由 SKIPMAX 改名，名实对齐）/ the counter anti wrap clamp bound
END_VAR

// 段 0｜沿检测无条件周期刷新（禁入分支）/ segment 0, the unconditional refresh
rtReset(CLK := bReset); // 复位沿 / the reset edge

// 段 1｜首扫初始化（R310）：环清零与指针复位（与复位沿同款块）/ segment 1, the first scan init, the same block as the reset edge
IF NOT _bInit THEN // 首扫一拍 / the first scan
    _bInit := TRUE; // 置首扫标志 / raise the flag
    FOR _nI := 0 TO 4095 DO // 固定界清环 / the fixed bound ring clear
        _aRing[_nI] := 0.0; // 槽清零 / clear the slot
    END_FOR
    _uWidx := 0; // 指针复位 / reset the index
    _nTick := 0; // 拍计数复位 / reset the tick count
END_IF

// 段 2｜复位沿作用域：清环 / 清指针与计数 / 清锁存（三项逐项声明）/ segment 2, the reset edge scope
IF rtReset.Q THEN // 复位沿 / the reset edge
    FOR _nI := 0 TO 4095 DO // 作用域一：固定界清环 / scope one, the fixed bound ring clear
        _aRing[_nI] := 0.0; // 槽清零 / clear the slot
    END_FOR
    _uWidx := 0; // 作用域二：清写指针 / scope two, clear the write index
    _nTick := 0; // 作用域二：清累计拍 / scope two, clear the tick count
    nSkipCnt := 0; // 作用域二：清拒收计数 / scope two, clear the skip count
    _bLatch := FALSE; // 作用域三：清域闸锁存（解除路径 = bReset 沿，R188）/ scope three, clear the latch
END_IF

// 段 3｜组态域闸（边界一）/ segment 3, the config gate
_nPer := UINT_TO_DINT(nPeriodTicks); // 升宽工作副本 / the widened work copy
IF (nPeriodTicks < 2) OR (nPeriodTicks > DL_PDC_PERMAX) // 周期域 / the period domain
OR (fForget < 0.0) OR (fForget > DL_PDC_FGTMAX) // 遗忘因子域（禁 1.0 无界累积）/ the forgetting domain
OR (fGain < 0.0) OR (fGain > 1.0) // 收敛增益域 / the gain domain
OR (fForget <> fForget) OR ((fForget - fForget) <> (fForget - fForget)) // 遗忘因子非有限 / a non finite forgetting
OR (fGain <> fGain) OR ((fGain - fGain) <> (fGain - fGain)) THEN // 增益非有限 / a non finite gain
    IF NOT _bLatch THEN // 未锁存才置位 / latch only while unlatched
        _bLatch := TRUE; // 置域闸锁存 / raise the latch
    END_IF
END_IF
bError := _bLatch; // 故障标志与锁存位同源（R191 名实双出口）/ the flag shares the latch

// 段 4｜内模逐拍正反馈累加（先读后写，边界二）/ segment 4, the internal model per tick, read then write
_bFin := (fErr = fErr) AND ((fErr - fErr) = (fErr - fErr)); // 误差有限双判据（R79）/ the error finiteness dual verdicts
IF bEnable AND (NOT _bLatch) AND _bFin THEN // 使能且域内且样本有限 / enabled, inside the domain, and finite
    fComp := -fGain * _aRing[_uWidx]; // 读上周期同相位存量取负前馈（写指针槽界已证 0..4095）/ the negative feedforward of the stored same phase error
    _aRing[_uWidx] := fErr + fForget * _aRing[_uWidx]; // 写本拍泄漏积分 / write the leaked integration
    _uWidx := _uWidx + 1; // 拍推进 / advance the tick
    IF UINT_TO_DINT(_uWidx) >= _nPer THEN // 按新周期回绕（比较式回绕，无 MOD 无移位）/ wrap by the period comparison
        _uWidx := 0; // 回绕到零 / wrap to zero
    END_IF
    IF _nTick < DL_PDC_CNTMAX THEN // 累计拍防回绕 / the tick wrap guard
        _nTick := _nTick + 1; // 累计推进 / advance the count
    END_IF
    bLearned := (_nTick >= DINT_TO_UDINT(_nPer)); // 环已填满一周期判定（标准转换函数）/ the filled verdict with a standard conversion
ELSIF (NOT _bFin) AND (NOT _bLatch) AND bEnable THEN // 非有限拒收拍（边界三）：环不写输出冻结 / a non finite tick, the ring untouched, the output frozen
    IF nSkipCnt < DL_PDC_CNTMAX THEN // 拒收计数防回绕 / the skip wrap guard
        nSkipCnt := nSkipCnt + 1; // 拒收计数推进 / advance the skip count
    END_IF
ELSE // 失能或域闸锁存：输出安全侧零（边界一）/ disabled or latched, the output safe zero
    fComp := 0.0; // 安全侧零 / the safe zero
    bLearned := FALSE; // 填满指示随失能清除 / the indicator cleared
END_IF
END_FUNCTION_BLOCK
